(* IEC 61131-3 sources: daoli-st-library/DL_MathData (part 27) *)

(* ---- FC_DL_TrimmedMeanCalc.st ---- *)
(*
  ==================================================================
  组件名 Component  : FC_DL_TrimmedMeanCalc
  分类   Category   : DL_MathData
  前缀   Naming     : FC_DL_ ｜ b/n/u/f/t/e/st 类型前缀制（R265）
  码位   Code ID    : 16#0001_0659 / 065A（故障级）
  版本   Version    : 1.0.0
  复杂度 Complexity  : 中
  功能   Purpose    : 双端截尾均值（稳健统计，抗野点污染的位置估计）：剔除非有限
                      样本后按升序索引对中段区间求均值。
  开源溯源 Origin    : 公开公式 clean-room，参考公开稳健统计教材的双端截尾均值
                      定义（分类与公式借鉴，零代码复制），本件实现、闸门与码位
                      100% 自有。
  许可证 License    : MIT
  参考   Reference  : IEC 61131-3:2013 §6.6 算术运算符；trimmed mean 公开统计定义
  平台   Platform   : 纯 IEC 61131-3（FOR / 四则 / 委托），三平台通用
  依赖   Depends    : FC_DL_SortIndexLReal（索引排序属主，本件委托排序，R140）
  分工声明 Split     : FC_DL_MeanAbsDevCalc（离散度）/ FC_DL_MedianAbsDev（稳健
                      离散度）/ FB_DL_MovingAverage（滑窗均值）互引；本件为双端
                      截尾均值（稳健位置估计），填位置量缺口（R216）。
  归属 Ownership     : 本件无 TYPE 声明；全部引脚为 IEC 标准原生类型。
                      委托件码位随其属主回传（R66）。
  ------------------------------------------------------------------
  边界 Boundary     :
                      一 非有限样本逐条剔除并计入局部 nNonFinite；nNonFinite 口径
                         **不外显**（R62-D7 定稿口径固化），剔除诊断请用
                         FC_DL_SignalStatistics；除子一律用剔除后的 nEff；
                      二 nCount 越域（< 1 或 > 256）或剔净后 nEff = 0 → 故障码
                         0659 早退（除子已证 ≥ 1 才进入均值段）；
                      三 uTrimLo + uTrimHi >= nEff → 组态码 065A 早退（禁把截尾
                         做成空集）；trim 以剔除后有效样本为基准（非入参计数）；
                      四 委托排序返回值与 bValid 由两个独立变量承接后合取
                         （R295 双承接）；委托码随属主回传（R66）；
                      五 均值区间 [uTrimLo, nEff−1−uTrimHi]，除子
                         (nEff − uTrimLo − uTrimHi) ≥ 1 由段 3 闸证明（禁除零）；
                      六 结果复检非有限 → 三件套兜底（R258）；
                      七 纯函数：无记忆量、无定时器、无边沿实例，每调用重算；
                      八 无全局、无外部变量、无物理地址、无指针。
  错误码 Codes      :
    16#0001_0659【故障级】有效样本数越域（nCount < 1 / > 256，或剔净后 nEff = 0）
    16#0001_065A【故障级】截尾组态非法（uTrimLo + uTrimHi >= nEff，截尾成空集）
  码位反证 Note     :
    0659 与 065A 不可合并：前者出口 nEff = 0（无任何有效样本），后者出口 nEff ≥ 1
    （有效样本存在但被截空），nEff 可由输出唯一还原场景（R90）；0659 合并
    「入参越域」与「剔净为空」的理由：两者出口组合完全同形（fMean = 0、nEff = 0、
    bValid = FALSE），按 R90 不另立。
  验收 Acceptance   :
    算法已证（脚本）：未跑 ｜ 编译器已证（三平台）：未跑
    V1 全同样本 + 任意 trim → 均值 = 该值
    V2 trim = 0/0 → 等价普通均值；V3 uTrimLo+uTrimHi = nEff → 码 065A 早退
    V4 nEff − trim = 1（只余 1 个）→ 均值 = 该样本
    V5 nCount = 0 → 码 0659；V6 nCount = 257 → 码 0659 早退
    V7 含 2 个 NaN → nEff 正确缩减（量化断言）
    V8 trim 单端不对称（lo = 2, hi = 0）→ 区间正确
  修订记录 Revision  :
    2026-11-21  v1.0.0  R63 首版（批 2 · 序号 4）
  ==================================================================
*)
FUNCTION FC_DL_TrimmedMeanCalc : BOOL
VAR_IN_OUT
    afSamples : ARRAY[0..255] OF LREAL; // 样本序列 [工程单位]，只读 / the sample series, read only
END_VAR
VAR_INPUT
    nCount  : DINT := 0;    // 有效样本数入参 [个]，合法域 1..256 / the sample count, legal from one to two hundred fifty six
    uTrimLo : USINT := 0;   // 低端截去个数 [个] / the count trimmed from the low end
    uTrimHi : USINT := 0;   // 高端截去个数 [个] / the count trimmed from the high end
END_VAR
VAR_OUTPUT
    fMean   : LREAL := 0.0; // 截尾均值 [工程单位] / the trimmed mean
    nEff    : DINT := 0;    // 参与均值样本数 [个]（剔除非有限后）/ the effective sample count after dropping non finite samples
    bValid  : BOOL := FALSE; // 结果可用 [-] / the result usable flag
    eErr    : UDINT := 16#0000_0000; // 错误码，0 = 正常 / the error code, zero is ok
    bError  : BOOL := FALSE; // 故障标志（故障级码同拍置位，R45 配对）/ the fault flag raised with a fault level code
END_VAR
VAR
    aVal      : ARRAY[0..255] OF LREAL; // 剔除非有限后的有效样本副本 [工程单位] / the finite sample copy
    aIdx      : ARRAY[0..255] OF DINT;  // 委托输出的排序索引排列 [下标] / the sorted permutation from the delegate
    k         : DINT := 0;    // 遍历索引 [下标] / the traversal index
    nNonFinite: DINT := 0;    // 剔除的非有限样本数 [个]（仅局部留档，不外显，R62-D7 口径；诊断请用 FC_DL_SignalStatistics）/ the dropped non finite count, local only and never exposed
    nCountUse : DINT := 0;    // 入参样本数接管量 [个] / the raw input count holder
    nTrim     : DINT := 0;    // 双端截去总数 [个]（升位防 USINT 和溢出）/ the total trimmed count widened before the sum
    nTrimLo   : DINT := 0;    // 低端截去数升位副本 [个] / the low trim count widened
    nTrimHi   : DINT := 0;    // 高端截去数升位副本 [个] / the high trim count widened
    nKeep     : DINT := 0;    // 参与均值样本数（除子）[个] / the kept sample count used as the divisor
    fSum      : LREAL := 0.0; // 区间样本和 [工程单位] / the interval sample sum
    fMeanUse  : LREAL := 0.0; // 均值工作副本 [工程单位] / the working mean copy
    bSortRet  : BOOL := FALSE; // 委托返回值承接量（独立承接，R295）/ the delegate return holder
    bSortValid: BOOL := FALSE; // 委托 bValid 承接量（独立承接，R295）/ the delegate valid holder
    uSortErr  : UDINT := 16#0000_0000; // 委托错误码承接量 [码] / the delegate error code holder
    bSortErr  : BOOL := FALSE; // 委托故障位承接量 / the delegate fault bit holder
    bSortOk   : BOOL := FALSE; // 返回值与可用位合取后的排序可用位 / the conjunction of the return value and the valid flag
END_VAR  // R64 结构补齐：VAR 段缺失的 END_VAR（门禁机械修复）
VAR CONSTANT
    DL_TMC_NMAX  : DINT := 256;      // 样本容量上界 [个]，与数组容量一致 / the capacity aligned with the array
    DL_TMC_ONE   : DINT := 1;        // 整型一常量 [个] / the integer one constant
    DL_TMC_ZERO  : DINT := 0;        // 整型零常量 [个] / the integer zero constant
END_VAR

// 段 1｜返回值与全部出口预置安全值（R45 四段式第一段）/ segment 1, the preset of the return and every outlet
FC_DL_TrimmedMeanCalc := FALSE; // 返回值预置假 / preset the return false
fMean := 0.0; // 均值预置零 [工程单位] / preset the mean zero
nEff := DL_TMC_ZERO; // 有效样本数预置零 [个] / preset the effective count zero
bValid := FALSE; // 可用标志预置假 / preset the validity false
eErr := 16#0000_0000; // 错误码预置正常 / preset the code to ok
bError := FALSE; // 故障标志预置假 / preset the error flag false
nNonFinite := DL_TMC_ZERO; // 剔除计数预置零 [个] / preset the dropped count zero
nCountUse := DL_TMC_ZERO; // 入参计数接管量预置零 [个] / preset the raw count holder zero
nTrim := DL_TMC_ZERO; // 截去总数预置零 [个] / preset the trimmed total zero
nTrimLo := DL_TMC_ZERO; // 低端截去数预置零 [个] / preset the low trim zero
nTrimHi := DL_TMC_ZERO; // 高端截去数预置零 [个] / preset the high trim zero
nKeep := DL_TMC_ZERO; // 除子预置零 [个] / preset the divisor zero
fSum := 0.0; // 区间和预置零 [工程单位] / preset the interval sum zero
fMeanUse := 0.0; // 均值工作副本预置零 [工程单位] / preset the working mean zero
bSortRet := FALSE; // 委托返回值承接量预置假 / preset the delegate return holder false
bSortValid := FALSE; // 委托可用位承接量预置假 / preset the delegate valid holder false
uSortErr := 16#0000_0000; // 委托码承接量预置零 [码] / preset the delegate code zero
bSortErr := FALSE; // 委托故障位承接量预置假 / preset the delegate fault holder false
bSortOk := FALSE; // 排序可用位预置假 / preset the sort usable bit false

// 段 2｜样本数域闸（边界二，早退禁除零）/ segment 2, the sample count domain gate
nCountUse := nCount; // 入参计数接管 [个] / take the raw count
IF (nCountUse < DL_TMC_ONE) OR (nCountUse > DL_TMC_NMAX) THEN // 计数越域 / the count is out of the domain
    eErr := 16#0001_0659; // 故障级：有效样本数越域 / fault grade, the effective sample count is out of the domain
    bError := TRUE; // 同拍置故障标志（R45 配对）/ raise the fault flag on the same scan
    bValid := FALSE; // 结果不可用 / the result is not usable
    RETURN; // 早退 / early return
END_IF

// 段 3｜非有限样本剔除（边界一：除子口径 = 剔除后有效样本数）/ segment 3, drop the non finite samples
FOR k := DL_TMC_ZERO TO nCountUse - DL_TMC_ONE DO // 有界遍历（上界已证 ≤ 256）/ the bounded traversal with a proven ceiling
    IF (afSamples[k] = afSamples[k]) AND ((afSamples[k] - afSamples[k]) = (afSamples[k] - afSamples[k])) THEN // 有限样本 / a finite sample
        aVal[nEff] := afSamples[k]; // 有限样本写入副本 [工程单位] / copy the finite sample
        nEff := nEff + DL_TMC_ONE; // 有效计数推进 [个] / advance the effective count
    ELSE // 非有限样本 / a non finite sample
        nNonFinite := nNonFinite + DL_TMC_ONE; // 剔除计数推进（仅局部留档，不外显）/ advance the dropped count, local only
    END_IF
END_FOR
IF nEff < DL_TMC_ONE THEN // 剔净后无有效样本（与段 2 同码，出口组合不可区分，R90）/ no sample remains after the drop
    eErr := 16#0001_0659; // 故障级：有效样本数越域（此处为剔净后为空）/ fault grade, the effective count is empty after the drop
    bError := TRUE; // 同拍置故障标志（R45 配对）/ raise the fault flag on the same scan
    bValid := FALSE; // 结果不可用 / the result is not usable
    RETURN; // 早退 / early return
END_IF

// 段 4｜截尾组态闸（边界三，trim 以 nEff 为基准；升位防 USINT 和回绕）/ segment 4, the trim configuration gate
nTrimLo := USINT_TO_DINT(uTrimLo); // 低端截去数升位 [个] / widen the low trim count
nTrimHi := USINT_TO_DINT(uTrimHi); // 高端截去数升位 [个] / widen the high trim count
nTrim := nTrimLo + nTrimHi; // 双端总数（DINT 域无回绕）[个] / the trimmed total in the widened domain
IF nTrim >= nEff THEN // 截尾成空集 / the trim leaves an empty set
    eErr := 16#0001_065A; // 故障级：截尾组态非法 / fault grade, the trim configuration is illegal
    bError := TRUE; // 同拍置故障标志（R45 配对）/ raise the fault flag on the same scan
    bValid := FALSE; // 结果不可用 / the result is not usable
    RETURN; // 早退，除子 nKeep 不可为零 / early return, the divisor can never reach zero
END_IF
nKeep := nEff - nTrim; // 参与均值样本数（除子）[个]，已证 ≥ 1 / the kept count, proven at least one

// 段 5｜委托索引排序（R140；返回值与可用位分承后合取，R295）/ segment 5, the delegated index sort
bSortRet := FC_DL_SortIndexLReal(afValues := aVal, nCount := nEff, aIdx => aIdx, bValid => bSortValid, eErr => uSortErr, bError => bSortErr); // 委托排序：两路各自承接 / delegate the sort into two distinct holders
bSortOk := bSortRet AND bSortValid; // 返回值与可用位合取（IEC 未规定两者的求值次序）/ conjoin the two signals since their evaluation order is unspecified
IF (NOT bSortOk) OR bSortErr THEN // 委托失败 / the delegate failed
    eErr := uSortErr; // 委托码回传（码随属主，R66）/ replay the delegate code
    bError := bSortErr; // 委托故障位回传 / replay the delegate fault bit
    bValid := FALSE; // 结果不可用 / the result is not usable
    RETURN; // 早退 / early return
END_IF

// 段 6｜区间求和（索引区间 [uTrimLo, nEff−1−uTrimHi]；除子 nKeep 已证 ≥ 1，边界五）/ segment 6, the interval sum over the trimmed range
FOR k := nTrimLo TO (nEff - DL_TMC_ONE) - nTrimHi DO // 有界遍历中段区间（区间端点已证合法）/ the bounded traversal over the kept range with proven endpoints
    fSum := fSum + aVal[aIdx[k]]; // 区间样本累加 [工程单位] / accumulate the kept samples
END_FOR
fMeanUse := fSum / DINT_TO_LREAL(nKeep); // 截尾均值 = 和 ÷ 参与数 [工程单位]，除子已证 ≥ 1 / the trimmed mean with the proven divisor

// 段 7｜结果复检兜底（三件套，R258）/ segment 7, the result recheck with the three part fallback
IF (fMeanUse <> fMeanUse) OR ((fMeanUse - fMeanUse) <> (fMeanUse - fMeanUse)) THEN // 结果非有限（理论上不可达，防御保留）/ a non finite result, unreachable by theory, kept as a defence
    fMean := 0.0; // 兜底安全值 [工程单位] / the bottom line safe value
    nEff := DL_TMC_ZERO; // 有效数清零（出口与故障场景同形）/ clear the effective count
    eErr := 16#0001_0659; // 故障级：结果非有限（与样本数越域同族一码，出口组合不可区分，R90）/ fault grade under the same family code
    bError := TRUE; // 置故障标志（R45 配对）/ raise the fault flag
    bValid := FALSE; // 结果不可用 / the result is not usable
    RETURN; // 早退 / early return
END_IF

// 段 8｜统一出口 / segment 8, the unified outlet
fMean := fMeanUse; // 均值出口 [工程单位] / the mean outlet
bValid := TRUE; // 结果可用 / the result is usable
FC_DL_TrimmedMeanCalc := TRUE; // 返回成功 / return success
END_FUNCTION

(* ---- FC_DL_TruncEx.st ---- *)
(*
    FC_DL_TruncEx —— 向零取整防御包装（DINT 范围钳位 + NaN 拦截）
    ------------------------------------------------------------------
    分类      : DL_MathData / Math-Round
    前缀      : FC_DL_
    版本      : 1.0.0
    溯源      : IEC 61131-3 标准语义的道莅防御性实现
                （内部委托平台内建函数，外围统一错误码/钳位/双语文档；
                  未复制任何闭源厂商源码，参考实现仅限 MIT/Apache 许可）
    平台      : 纯 IEC 61131-3，CODESYS / TwinCAT / InoProShop 通用
    作者      : 道莅代码库 · PLC编程专家（R15）
    ------------------------------------------------------------------
    功能说明  : 向零取整（委托内建 TRUNC），如 1.9 得 1、-1.9 得 -1。
                NaN 输入拦截返回 0 并置 16#0001_018B；结果超 DINT 范围
                [-2147483648, 2147483647] 时钳位到对应边界并置 16#0001_0259
                （钳位值非真实取整，bValid=FALSE；无穷输入被范围闸自然
                拦截）。先做范围闸再调 TRUNC，保证内建转换永不溢出。
    错误码    : 0000 正常 / 16#0001_018B 入参越界（NaN 已归零） / 16#0001_0259 上溢下溢（已钳位到 DINT 边界）
    修订记录  : 2026-11-16 v1.0.0 首次入库（R15）
*)
FUNCTION FC_DL_TruncEx : DINT
VAR_INPUT
    lrIn : LREAL; // 输入实数 [无量纲]，任意有限值或 NaN/无穷 / input real value [dimensionless], any finite value or NaN/inf
END_VAR
VAR_OUTPUT
    eErr : UDINT; // 错误码，0=正常，1=入参越界，2=上溢下溢 / error id, 0=ok, 1=input out of domain, 2=overflow or underflow
    bError   : BOOL; // 是否出错，eErr 非 0 时为 TRUE / error flag, TRUE when eErr is nonzero
    bValid   : BOOL; // 输出是否有效可用，钳位降级时为 FALSE / output valid, FALSE for clamped degraded results
END_VAR
VAR CONSTANT
    DL_TR_HI : LREAL := 2147483648.0; // DINT 上溢闸 [无量纲]，入参达到即超界 / DINT upper overflow gate [dimensionless]
    DL_TR_LO : LREAL := -2147483649.0; // DINT 下溢闸 [无量纲]，入参达到即超界 / DINT lower overflow gate [dimensionless]
END_VAR

// 段 1｜返回值与错误状态预置，任何早退路径不留脏码 / segment 1, preset return value and error states
FC_DL_TruncEx := 0; // 返回值预置安全值 0 / preset return to safe value 0
eErr      := 16#0000_0000; // 错误码预置正常 / preset error id to ok
bError        := FALSE; // 错误标志预置无错 / preset error flag to FALSE
bValid        := TRUE; // 有效标志预置可用 / preset valid flag to TRUE

// 段 2｜NaN 拦截：自不等判据，归零早退，不进内核 / segment 2, NaN interception by self-inequality, zeroed early exit
IF lrIn <> lrIn THEN
    eErr := 16#0001_018B; // 信息级：输入 NaN，已归零 / informational, NaN input, zeroed
    bError   := TRUE; // 置错误标志 / raise error flag
    bValid   := FALSE; // 输出不可用 / output invalid
    RETURN; // 返回预置安全值 0 / return preset safe value 0
END_IF

// 段 3｜DINT 范围闸：先判后转换，保证内建 TRUNC 永不溢出（无穷输入同样命中闸） / segment 3, DINT range gate, decide before conversion so built-in TRUNC never overflows, infinity hits the gate too
IF lrIn >= DL_TR_HI THEN
    FC_DL_TruncEx := 2147483647; // 上溢钳位到 DINT 上界 / overflow clamped to the DINT upper bound
    eErr      := 16#0001_0259; // 上溢码 / overflow code
    bError        := TRUE; // 置错误标志 / raise error flag
    bValid        := FALSE; // 钳位值非真实取整 / clamped value is not the true truncation
    RETURN;
ELSIF lrIn <= DL_TR_LO THEN
    FC_DL_TruncEx := -2147483648; // 下溢钳位到 DINT 下界 / underflow clamped to the DINT lower bound
    eErr      := 16#0001_0259; // 下溢码 / underflow code
    bError        := TRUE; // 置错误标志 / raise error flag
    bValid        := FALSE; // 钳位值非真实取整 / clamped value is not the true truncation
    RETURN;
END_IF

// 段 4｜域内委托内建 TRUNC（向零取整） / segment 4, in-domain delegation to built-in TRUNC, rounding toward zero
FC_DL_TruncEx := TRUNC(lrIn); // 委托内建 TRUNC 内核，不自实现取整内核 / delegate to built-in TRUNC kernel

// 段 5｜结果复检兜底（防御纵深，正常路径不可达） / segment 5, result recheck as defense in depth
IF (FC_DL_TruncEx <> FC_DL_TruncEx) OR (FC_DL_TruncEx > 2147483647) OR (FC_DL_TruncEx < -2147483648) THEN
    FC_DL_TruncEx := 0; // 兜底安全值 / bottom-line safe value
    IF eErr = 16#0000_0000 THEN
        eErr := 16#0001_018B; // 首事件优先置码 / first-event priority code
        bError   := TRUE; // 置错误标志 / raise error flag
        bValid   := FALSE; // 输出不可用 / output invalid
    END_IF
END_IF
END_FUNCTION

(* ---- FC_DL_TruncToMultipleInt.st ---- *)
(*==============================================================================
 * 组件名称 : FC_DL_TruncToMultipleInt ｜ 子库 : DL_MathData ｜ v1.0.0 ｜ 2026-11-23
 * 平台     : CODESYS 3.5 / TwinCAT 3 / InoProShop / Machine Expert（纯 IEC，无厂商库）
 * 功能简介 : 整数向零截断到 nMultiple 的倍数（丢弃不足一个倍数的余量，
 *            符号随被除数）。纯整数算术实现：整除（ST 中 DIV 对整数
 *            向零截断）后回乘，即得截断对齐结果。
 * 契约     : 返回向零截断结果；nMultiple <= 0 恒返回 0；
 *            纯函数无状态、同输入同输出。
 * 依赖     : 无 DL_ 内部依赖（本批自足实现）
 * 红线自检 : R1 零全局 R2 零%I/%Q R3 纯IEC R4 非法倍数返 0（防除零）
 *            R5 双语注释 R6 N/A（无状态机） R7 N/A（无定时器实例）
 * 修订历史 : 2026-11-23 R78-B1 对齐取整族模板派生首版
 *============================================================================*)
FUNCTION FC_DL_TruncToMultipleInt : DINT
VAR_INPUT
    nValue : DINT;          // 输入整数 / Input integer value
    nMultiple : DINT;       // 对齐倍数，须 > 0 / Alignment multiple, must be > 0
END_VAR
IF nMultiple <= 0 THEN
    FC_DL_TruncToMultipleInt := 0;      // 非法倍数返 0 / Invalid multiple returns 0
    RETURN;
END_IF
FC_DL_TruncToMultipleInt := (nValue / nMultiple) * nMultiple;   // 整除截断回乘 / Truncate by integer division and remultiply
END_FUNCTION

(* ---- FC_DL_UdintToBcd.st ---- *)
(*
    FC_DL_UdintToBcd —— UDINT 到 8 位十进制 BCD 码饱和防御转换
    ------------------------------------------------------------------
    分类      : DL_MathData / Convert
    前缀      : FC_DL_
    版本      : 1.0.0
    溯源      : IEC 61131-3 标准语义的道莅防御性实现
                （内部委托平台内建函数，外围统一错误码/钳位/双语文档；
                  未复制任何闭源厂商源码，参考实现仅限 MIT/Apache 许可）
    平台      : 纯 IEC 61131-3，CODESYS / TwinCAT / InoProShop 通用
    作者      : 道莅代码库 · PLC编程专家（R16）
    ------------------------------------------------------------------
    功能说明  : 将十进制值 nIn（0..99999999）防御性转换为 8 位十进制 BCD 码并返回；
                nIn 超出 99999999 时饱和输出 BCD 码 16#99999999，置信息级 16#0001_01D2
                （与 R9 FC_DL_WordToBcd 的 9999 饱和口径一致，域扩大 4 位）；
                钳位方向：仅上界单侧饱和至 16#99999999；
                域内按除 10 取余逐位拼装半字节：除子为常量 10，编译期恒非零，
                满足除法前判除子非零红线；8 次整除后余数归零，无溢出路径；
                纯整数域输入不存在 NaN/±INF 非有限态，故本组件无故障级路径；
                信息级码属正常防御：bError=FALSE、bValid=TRUE，输出饱和后防御值。
    错误码    : 16#0001_01D2 输入超 99999999，已饱和至 BCD 16#99999999——信息级，正常防御
                16#0001_01D3 预留禁用（信息级，不得挪用）
                16#0001_02A9 预留禁用（故障级，不得挪用）
                16#0001_02AA 预留禁用（故障级，不得挪用）
                16#0001_02AB 预留禁用（故障级，不得挪用）
    状态机    : R6 标注 N/A —— 本组件为纯函数无顺序状态机，无 CASE 可写，非法状态不可能出现，故以本节说明替代 ELSE 兜底
    修订记录  : 2026-11-16 v1.0.0 首次入库（R16）
*)
FUNCTION FC_DL_UdintToBcd : UDINT
VAR_INPUT
    nIn : UDINT; // 十进制值 [0..99999999] / decimal value, 0..99999999
END_VAR
VAR_OUTPUT
    eErr   : UDINT; // 错误码，0=正常 / error id, 0=ok
    bError : BOOL;  // 是否出错，eErr 非 0 时为 TRUE / error flag, TRUE when eErr is nonzero
    bValid : BOOL;  // 输出是否有效可用 / output valid flag
END_VAR
VAR CONSTANT
    DL_BCD8_MAX    : UDINT := 99999999;    // 8 位 BCD 十进制域上界 [无量纲] / 8-digit BCD decimal domain upper bound
    DL_BCD8_SAT    : UDINT := 16#99999999; // 8 位 BCD 饱和输出码（每位半字节 9） [BCD 位] / 8-digit BCD saturating output code (nibble 9 each)
    DL_BCD_NIB_CNT : INT   := 8;           // UDINT 32 位容器 BCD 半字节总数 [个] / total BCD nibble count of 32-bit UDINT container
    DL_DEC_BASE    : UDINT := 10;          // 十进制除法基（编译期常量，恒非零） [基数] / decimal division base (compile-time constant, never zero)
END_VAR
VAR
    i      : INT;   // 半字节循环索引 [个] / nibble loop index
    uDigit : UDINT; // 当前十进制位值（0~9） [位] / current decimal digit value (0~9)
    uTmp   : UDINT; // 剩余待转换商 [无量纲] / remaining quotient to convert
END_VAR

// 段 1｜返回值与错误状态预置 / segment 1, preset return value and error status
FC_DL_UdintToBcd := 0; // 故障缺省返回 0 [BCD 位] / fault default returns 0
eErr   := 0;     // 预置无错误 / preset no error
bError := FALSE; // 预置无故障（整数域无故障态） / preset no fault (no fault states in integer domain)
bValid := FALSE; // 预置无效，通过饱和判定后置位 / preset invalid, set TRUE after saturation check

// 段 2｜上界单侧饱和钳位 / segment 2, upper-bound saturating clamp
IF nIn > DL_BCD8_MAX THEN
    FC_DL_UdintToBcd := DL_BCD8_SAT; // 饱和输出 BCD 16#99999999（与 R9 WordToBcd 口径一致，域扩大 4 位） / saturate to BCD 16#99999999 (aligned with R9 WordToBcd policy, domain widened by 4 digits)
    eErr := 16#0001_01D2;            // 信息级：超上界已饱和 / info level: above upper bound, saturated
    bError := FALSE;                 // 信息级饱和不置故障 / info-level saturation never raises fault
    bValid := TRUE;                  // 饱和输出有效可用 / saturated output is valid
    RETURN;                          // 立即返回 / immediate return
END_IF

// 段 3｜除 10 取余逐位拼装主体计算（末段） / segment 3, divide-by-10 remainder digit assembly main conversion (final)
uTmp := nIn; // 商初始化为输入值 / initialize quotient with input
FOR i := 0 TO DL_BCD_NIB_CNT - 1 DO
    uDigit := uTmp MOD DL_DEC_BASE;       // 除 10 取余得当前十进制位（除子常量 10 恒非零） / modulo 10 for current digit (constant divisor 10, never zero)
    FC_DL_UdintToBcd := FC_DL_UdintToBcd OR SHL(uDigit, 4 * i); // 拼装第 i 个 BCD 半字节（SHL 移位量 4*i ≤ 28 安全） / assemble i-th BCD nibble (shift 4*i <= 28, safe)
    uTmp := uTmp / DL_DEC_BASE;           // 整除 10 前进到下一位（除子常量 10 恒非零） / integer-divide by 10 to next digit (constant divisor 10, never zero)
END_FOR
bError := FALSE; // 域内转换无故障 / in-domain conversion, no fault
bValid := TRUE;  // 输出有效可用 / output valid
END_FUNCTION

(* ---- FC_DL_UdintToDintChk.st ---- *)
(*
    FC_DL_UdintToDintChk —— UDINT 到 DINT 越界钳位防御转换
    ------------------------------------------------------------------
    分类      : DL_MathData / Convert
    前缀      : FC_DL_
    版本      : 1.0.0
    溯源      : IEC 61131-3 标准语义的道莅防御性实现
                （内部委托平台内建函数，外围统一错误码/钳位/双语文档；
                  未复制任何闭源厂商源码，参考实现仅限 MIT/Apache 许可）
    平台      : 纯 IEC 61131-3，CODESYS / TwinCAT / InoProShop 通用
    作者      : 道莅代码库 · PLC编程专家（R16）
    ------------------------------------------------------------------
    功能说明  : 将 UDINT 输入防御性转换为 DINT 并作为返回值输出；
                uIn 超出 DINT 上界 2147483647 时钳位至上界，置信息级 16#0001_01CC；
                钳位方向：仅上界单侧饱和（UDINT 无负值，下界 0 天然落在 DINT 域内无需钳位）；
                纯整数域输入不存在 NaN/±INF 非有限态，亦无除法运算，故本组件无故障级路径；
                域内转换委托平台内建 UDINT_TO_DINT 语义，不重实现数学内核；
                信息级码属正常防御：bError=FALSE、bValid=TRUE，输出钳位后防御值。
    错误码    : 16#0001_01CC 输入超 DINT 上界，已钳位至 2147483647——信息级，正常防御
                16#0001_01CD 预留禁用（信息级，不得挪用）
                16#0001_02A0 预留禁用（故障级，不得挪用）
                16#0001_02A1 预留禁用（故障级，不得挪用）
                16#0001_02A2 预留禁用（故障级，不得挪用）
    状态机    : R6 标注 N/A —— 本组件为纯函数无顺序状态机，无 CASE 可写，非法状态不可能出现，故以本节说明替代 ELSE 兜底
    修订记录  : 2026-11-16 v1.0.0 首次入库（R16）
*)
FUNCTION FC_DL_UdintToDintChk : DINT
VAR_INPUT
    uIn : UDINT; // 待转换输入 [无量纲] / input value to convert
END_VAR
VAR_OUTPUT
    eErr   : UDINT; // 错误码，0=正常 / error id, 0=ok
    bError : BOOL;  // 是否出错，eErr 非 0 时为 TRUE / error flag, TRUE when eErr is nonzero
    bValid : BOOL;  // 输出是否有效可用 / output valid flag
END_VAR
VAR CONSTANT
    DL_DINT32_MAX : UDINT := 2147483647; // DINT 域上界 2147483647 [无量纲] / DINT upper bound 2147483647
END_VAR

// 段 1｜返回值与错误状态预置 / segment 1, preset return value and error status
FC_DL_UdintToDintChk := 0; // 故障缺省返回 0 [无量纲] / fault default returns 0
eErr   := 0;     // 预置无错误 / preset no error
bError := FALSE; // 预置无故障（整数域无故障态） / preset no fault (no fault states in integer domain)
bValid := FALSE; // 预置无效，通过钳位判定后置位 / preset invalid, set TRUE after clamp check

// 段 2｜上界单侧饱和钳位与主体转换（末段） / segment 2, upper-bound saturating clamp and main conversion (final)
IF uIn > DL_DINT32_MAX THEN
    FC_DL_UdintToDintChk := DL_DINT32_MAX; // 正向钳位至 DINT 上界 2147483647 / clamp to DINT upper bound 2147483647
    eErr := 16#0001_01CC;                  // 信息级：超上界已钳位 / info level: above upper bound, clamped
ELSE
    FC_DL_UdintToDintChk := UDINT_TO_DINT(uIn); // 域内委托平台内建 _TO_ 转换语义 / in-domain delegate to built-in _TO_ conversion
    eErr := 0; // 域内无错误 / in-domain, no error
END_IF
bValid := TRUE; // 域内或钳位输出均有效可用 / in-domain or clamped output is valid
END_FUNCTION

(* ---- FC_DL_UdintToLintChk.st ---- *)
(*
    FC_DL_UdintToLintChk —— UDINT 到 LINT 升位验真
    ------------------------------------------------------------------
    分类      : DL_MathData / Convert
    前缀      : FC_DL_
    版本      : 1.0.0
    溯源      : IEC 61131-3 标准语义的道莅防御性实现（UDINT 32 位无符号 → LINT 64 位有符号）；
                委托平台内建 UDINT_TO_LINT 完成升位，本件不重实现数学内核；
                round-trip 验真判据、复核开关、错误分级与码位 100% 自有；
                clean-room 重写，未复制任何闭源厂商源码，参考实现仅限 MIT/Apache 许可
    平台      : 纯 IEC 61131-3，CODESYS V3.5+ / TwinCAT 3 / InoProShop 通用
    作者      : 道莅代码库 · PLC编程专家（R20）
    ------------------------------------------------------------------
    功能说明  : UDINT 到 LINT 在数学上恒无损（32 位无符号域完全落在 64 位有符号域内），
                但平台实现常见两种路径：直接零扩展（正确），或经 32 位有符号中间量再升位
                （错误：≥ 2^31 的值被符号扩展成负数）。后者在 DINT 中转站写法里反复出现，
                且编译期无告警、运行期只在超过 2147483647 时才显形，属隐蔽缺陷。
                本件的价值就是把这个隐性错误变成可判定的显式故障：
                核心防御：① round-trip 验真——把结果 LINT_TO_UDINT 反算回去，
                   与输入逐位相等才算无损；不等即判平台符号扩展错误（故障级）；
                ② 验真是判定式而非猜测式：只依赖 IEC 标准往返转换，不依赖任何平台内建语义；
                ③ bCheckEveryCall = FALSE 时跳过复核以降开销，但发信息级说明
                   「本拍未验真」，让审计侧知道该批数据没有复核保护；
                ④ 反算本身也在域内（LINT 结果必为 0~4294967295，若平台已错则反算必然不等），
                   不存在二次溢出风险。
                职责边界：有符号域内饱和归 FC_DL_LintToDintSat，双向无符号落地归
                FC_DL_LintToUdintSat；本件只承担「升位是否真正无损」的验真职责。
    编译门槛  : 主路径依赖平台内建 UDINT_TO_LINT 与 LINT_TO_UDINT，均为 IEC 61131-3
                标准转换函数，三平台标准库均提供，无厂商方言。
    错误码    : 16#0001_0414 调用方关闭逐次复核（bCheckEveryCall = FALSE），本拍未验真——信息级，值仍可用
                16#0001_0415 预留禁用（信息级，不得挪用）
                16#0001_033C round-trip 验真失败，平台把中间量经 32 位有符号路径符号扩展——故障级，bValid = FALSE
                16#0001_033D 预留（故障级，不得挪用）
                16#0001_033E 预留禁用（故障级，不得挪用）
    码位总账  : 16#0001_0414 用 / 16#0001_0415 预留 ｜ 16#0001_033C 用 / 16#0001_033D 预留 / 16#0001_033E 预留
    状态机    : R6 标注 N/A —— 本组件为纯函数无顺序状态机，无 CASE 可写，非法状态不可能出现
    采样约定  : 本件无定时器、无沿检测、无状态；单拍纯计算，结论与任务周期无关。
                复核开关是引脚量而非内部锁存，调用方可按数据重要性逐调用切换。
    修订记录  : 2026-11-16 v1.0.0 首次入库（R20）
*)
FUNCTION FC_DL_UdintToLintChk : LINT
VAR_INPUT
    uIn              : UDINT;                // 输入值 [无量纲]，全域 0~4294967295 / input value [dimensionless], full UDINT domain
    bCheckEveryCall  : BOOL := TRUE;          // TRUE = 每次调用都做 round-trip 复核 / TRUE performs the round-trip check on every call
END_VAR
VAR_OUTPUT
    eErr             : UDINT;                 // 错误码，0=正常 / error id, 0=ok
    bError           : BOOL;                  // 故障标志，eErr 为故障级时 TRUE / error flag, TRUE on fault-level eErr
    bValid           : BOOL;                  // 返回值是否可用（验真失败为 FALSE）/ return usable, FALSE when the round trip failed
    bRoundTripFail   : BOOL;                  // round-trip 复核失败标志 / round-trip check failed flag
END_VAR
VAR CONSTANT
    DL_UDINT_MAX     : UDINT := 16#FFFF_FFFF; // UDINT 上限值，域上限登记（类型本身即保证无需显式比较）[无量纲] / the UDINT maximum, registered domain top [dimensionless]
    DL_LINT_ZERO     : LINT := 0;             // 有符号零常量，避免裸字面量 [无量纲] / signed zero constant [dimensionless]
END_VAR
VAR
    liOut            : LINT;                  // 升位结果中间量 [无量纲] / widened result intermediate [dimensionless]
    uBack            : UDINT;                 // 反算回无符号的复核值 [无量纲] / back-converted value used by the check [dimensionless]
END_VAR

// 段 1｜返回值与错误状态预置 / segment 1, preset return value and error status
FC_DL_UdintToLintChk := DL_LINT_ZERO;         // 故障缺省返回 0 [无量纲] / fault default returns zero [dimensionless]
eErr := 0;                                    // 预置无错误 / preset no error
bError := FALSE;                              // 预置无故障 / preset no fault
bValid := FALSE;                              // 预置不可用，通过闸门后置位 / preset invalid, set TRUE after the gates
bRoundTripFail := FALSE;                      // 预置未失败 / preset no failure
liOut := DL_LINT_ZERO;                        // 中间量清零 / clear the intermediate

// 段 2｜主体：域内升位委托平台内建（数学上恒无损）/ segment 2, widen through the built-in, mathematically lossless
liOut := UDINT_TO_LINT(uIn);                  // 32 位无符号升 64 位有符号 [无量纲] / widen 32-bit unsigned into 64-bit signed [dimensionless]

// 段 3｜复核开关闸：关闭复核只发信息级，绝不伪装成已验真 / segment 3, check switch gate
IF NOT bCheckEveryCall THEN
    eErr := 16#0001_0414;                     // 信息级：本拍未验真，值仍可用 / info level, unchecked this cycle, still usable
    FC_DL_UdintToLintChk := liOut;            // 发布未复核的结果 / publish the unchecked result
    bValid := TRUE;                           // 未复核不等于不可用 / unchecked does not mean unusable
    RETURN;                                   // 出口 / exit
END_IF

// 段 4｜round-trip 验真：反算回去必须逐位相等 / segment 4, round-trip verification
uBack := LINT_TO_UDINT(liOut);                // 反算回无符号域 [无量纲] / convert back into the unsigned domain [dimensionless]
IF uBack <> uIn THEN
    bRoundTripFail := TRUE;                   // 标记验真失败 / flag the failed verification
    eErr := 16#0001_033C;                     // 故障级：平台符号扩展错误 / fault level, the platform sign-extended the value
    bError := TRUE;                           // 置故障标志 / raise the error flag
    bValid := FALSE;                          // 返回值不可用于后续运算 / the value must not enter later arithmetic
    FC_DL_UdintToLintChk := liOut;            // 仍发布结果供 HMI 对比观察 / still publish the value so HMI can compare it
    RETURN;                                   // 出口 / exit
END_IF

// 段 5｜发布验真通过的结果 / segment 5, publish the verified result
FC_DL_UdintToLintChk := liOut;                // 输出升位结果 [无量纲] / publish the widened result [dimensionless]
bValid := TRUE;                               // 验真通过即可用 / verified values are usable
END_FUNCTION

(* ---- FC_DL_UdintToRealChk.st ---- *)
(*
    FC_DL_UdintToRealChk —— UDINT 到 REAL 精度告警转换
    ------------------------------------------------------------------
    分类      : DL_MathData / Convert
    前缀      : FC_DL_
    版本      : 1.0.0
    溯源      : IEC 61131-3 标准语义的道莅防御性实现
                （接口语义由 IEC 61131-3 定义，内部委托平台内建 UDINT_TO_REAL，
                  外围统一错误码 / 钳位 / 双语文档；clean-room 重写，
                  未复制任何闭源厂商源码，参考实现仅限 MIT/Apache 许可）
    平台      : 纯 IEC 61131-3，CODESYS / TwinCAT / InoProShop 通用
    作者      : 道莅代码库 · PLC编程专家（R17）
    ------------------------------------------------------------------
    功能说明  : 将 UDINT 防御性转换为 REAL 并作为返回值输出，转换委托平台内建 UDINT_TO_REAL；
                nIn 超过 2^24（16777216，REAL 尾数 24 位可精确表示的整数上界）时，
                值照常转换输出，仅置信息级 16#0001_01FE 提示低位精度损失（bError=FALSE、bValid=TRUE）；
                负值分支结构性不存在（UDINT 为无符号类型，由类型系统保证），故无下界比较；
                本件只对 REAL 目标域立项：UDINT 全域 ≤ 2^32 远小于 2^53，转 LREAL 恒无损，
                故不设 UDINT 到 LREAL 的告警件（该结论在此声明，后续轮次不得重复立项）；
                钳位方向：无钳位（信息级仅记录，转换结果为最接近的可表值）。
    错误码    : 16#0001_01FE nIn 超 2^24 精度极限，转换值低位可能失真——信息级，正常防御
                16#0001_01FF 预留禁用（信息级，不得挪用）
                16#0001_02EB 预留禁用（故障级，不得挪用）
                16#0001_02EC 预留禁用（故障级，不得挪用）
                16#0001_02ED 预留禁用（故障级，不得挪用）
    状态机    : R6 标注 N/A —— 本组件为纯函数无顺序状态机，无 CASE 可写，非法状态不可能出现，故以本节说明替代 ELSE 兜底
    修订记录  : 2026-11-16 v1.0.0 首次入库（R17）
*)
FUNCTION FC_DL_UdintToRealChk : REAL
VAR_INPUT
    nIn : UDINT; // 待转换无符号整数值，建议域 0 ~ 4294967295 [无量纲] / unsigned integer to convert, suggested domain 0 .. 4294967295 [dimensionless]
END_VAR
VAR_OUTPUT
    eErr   : UDINT; // 错误码，0=正常 / error id, 0=ok
    bError : BOOL;  // 是否出错，eErr 非 0 时为 TRUE / error flag, TRUE when eErr is nonzero
    bValid : BOOL;  // 输出是否有效可用 / output valid flag
END_VAR
VAR CONSTANT
    DL_F24_MAX_U : UDINT := 16777216; // REAL 尾数 24 位可精确表示的无符号整数上界 2^24 [无量纲] / 2^24 exact-integer bound of REAL's 24-bit significand [dimensionless]
    DL_REAL_ZERO : REAL  := 0.0;      // 返回值预置零（本件无故障路径，仅作预置约定） [无量纲] / preset zero, no fault path in this component [dimensionless]
END_VAR

// 段 1｜返回值与错误状态预置 / segment 1, preset return value and error status
FC_DL_UdintToRealChk := DL_REAL_ZERO; // 预置 0.0（本件无故障级路径，仅作预置约定） [无量纲] / preset 0.0, no fault-level path in this component [dimensionless]
eErr   := 0;     // 预置无错误 / preset no error
bError := FALSE; // 预置无故障（本件无故障级路径） / preset no fault, no fault-level path here
bValid := FALSE; // 预置输出无效，通过精度判定后置位 / preset invalid, set TRUE after the precision check

// 段 2｜24 位尾数精度极限判定与主体转换（末段） / segment 2, 24-bit significand precision check and main conversion (final)
FC_DL_UdintToRealChk := UDINT_TO_REAL(nIn); // 值照常转换（委托平台内建转换语义），本件只告警不钳位 [无量纲] / convert as-is via the built-in conversion, this component warns but never clamps [dimensionless]
IF nIn > DL_F24_MAX_U THEN // 无符号类型仅需上界单侧比较，负值分支由类型系统结构性排除 [无量纲] / unsigned type only needs the upper-bound test, negative branch excluded by the type system [dimensionless]
    eErr := 16#0001_01FE; // 信息级：超 2^24 精度极限，低位可能失真，仅记录不钳位 / info level: beyond the 2^24 precision limit, low bits may lose accuracy, recorded only
ELSE
    eErr := 0;            // 精度域内无告警 / within the precision domain, no notice
END_IF
bError := FALSE; // 信息级精度告警不置故障 / info-level precision notice never raises fault
bValid := TRUE;  // 域内或精度告警输出均有效可用 / in-domain or precision-noticed output is valid
END_FUNCTION

(* ---- FC_DL_UdintToStringTrim.st ---- *)
(*
    FC_DL_UdintToStringTrim —— UDINT 到定宽十进制字段（右对齐）的防御字符串化
    ------------------------------------------------------------------
    分类      : DL_MathData / Convert
    前缀      : FC_DL_
    版本      : 1.0.0
    溯源      : IEC 61131-3 标准语义的道莅防御性实现（UDINT → STRING 定宽右对齐补位，
                委托平台内建 UDINT_TO_STRING 与标准串函数 LEN / LEFT / CONCAT；
                补位、四步截断样板、目标宽度闸、错误分级与码位 100% 自有；
                clean-room 编写，未复制任何闭源厂商源码）
    平台      : 纯 IEC 61131-3，CODESYS 3.5 / TwinCAT 3 / InoProShop / Machine Expert 通用
    作者      : 道莅代码库 · PLC编程专家（R69 构建轮 · 批 1 · N3）
    ------------------------------------------------------------------
    功能说明  : R22 定宽字段族的无符号补口。库内已有 FC_DL_DintToStringTrim（有符号，
                去前导空格左对齐）与 FC_DL_LrealToStringTrim（浮点）——本件补 UDINT
                方向，且语义与有符号版**异构**，不可互相替代：
                ① 有符号版做「修剪」（去掉平台补的前导空格后左对齐）；
                   本件做「定宽右对齐」（按目标宽度左补空格，供报表 / 报文定宽字段）。
                ② 上界语义异构：DINT 上界 2147483647 为 10 位数，UDINT 上界
                   4294967295 为 10 位数但**多一个符号位宽**——若把 UDINT 值先转 DINT
                   （现场常见写法），大于 2147483647 的值会翻成负数并输出「-294967296」
                   ！本件全程在 UDINT 域内字符串化，禁止任何有符号中转（R55/R56 口径：
                   浮点 / 有符号 → 无符号必须双分支显式，此处根本不做中转）。
                ③ 目标宽度 uFieldWidth 域 1..32：0 宽度无意义（故障级）；超 32 亦为故障级
                   ——补位源是 32 字符空格常量，宽度超过补位源时 LEFT 会静默返回全长，
                   表现为「字段比要求窄」，故必须在域闸挡住而不得靠钳位；
                   宽度小于实际位数且 bAllowTrunc = FALSE 时返回空串并报故障级，
                   绝不返回半截数值（把 4294967295 写成 429 上位机会当真数据）。
                补位实现：用常量空格串 + LEFT 取 nPad 个 + CONCAT 前缀，禁 WHILE 拼串
                （拼串随长度平方级增长，且串函数异常时会死循环）。
    错误码    : 16#0001_04F8 已按目标宽度左补空格（bPadded 可查）—— 信息级，值可用
                16#0001_04F9 发生截断且 bAllowTrunc = TRUE（bTruncated 可查）—— 信息级，值可用
                16#0001_03FA 目标宽度非法（uFieldWidth = 0）—— 故障级，返回空串
                16#0001_03FB 需要截断但 bAllowTrunc = FALSE —— 故障级，返回空串
    码位总账  : 16#0001_03FA / 03FB 用 ｜ 16#0001_04F8 / 04F9 用
    状态机    : R6 标注 N/A —— 纯函数无顺序状态机，无 CASE 可写，非法状态不可能出现
    采样约定  : 无定时器 / 无沿检测 / 无跨周期状态，结论与任务周期无关
    修订记录  : 2026-11-22 v1.0.0 首次入库（R69 构建轮 · 批 1 · N3）
*)
FUNCTION FC_DL_UdintToStringTrim : STRING(255)
VAR_INPUT
    uIn          : UDINT;                      // 待字符串化的无符号值 [无量纲]，全域 0..4294967295 / unsigned value, full UDINT domain
    uFieldWidth  : USINT := 10;                // 定宽字段宽度 [字符]，域 1..32 / fixed field width [characters], 1 to 32
    bAllowTrunc  : BOOL := FALSE;              // TRUE = 允许截断；FALSE = 需截断即故障 / TRUE allows truncation
END_VAR
VAR_OUTPUT
    eErr         : UDINT;                      // 错误码，0 = 正常 / error id, 0 = ok
    bError       : BOOL;                       // 故障标志，故障级码时为 TRUE / error flag, TRUE on fault level
    bValid       : BOOL;                       // 返回值是否可用（故障级为 FALSE）/ return usable, FALSE on fault level
    bPadded      : BOOL;                       // 本次做了左补空格 / left padding happened
    bTruncated   : BOOL;                       // 本次发生截断 / truncation happened
END_VAR
VAR CONSTANT
    DL_US_CAP    : INT := 255;                 // STRING 型长度上限 [字符]（R49 口径）/ STRING capacity [characters]
    DL_US_W_MIN  : USINT := 1;                 // 目标宽度下限 [字符] / field width floor [characters]
    DL_US_W_MAX  : INT := 32;                  // 目标宽度上限 [字符]，等于补位源空格串长度（超此宽度补位不可信）/ width ceiling [characters]
    DL_US_BLANKS : STRING(32) := '                                ';  // 32 个空格常量，补位源 [字符] / 32 blanks, the padding source
    DL_US_EMPTY  : STRING(1) := '';            // 空串常量，故障缺省返回 / empty string returned on faults
    DL_US_ZERO   : INT := 0;                   // 整型零常量，避免裸字面量 [字符] / integer zero constant
END_VAR
VAR
    sRaw         : STRING(255);                // 内建字符串化原始结果 / raw result of the built-in conversion
    sPad         : STRING(32);                 // 左补空格串 / left padding string
    sOut         : STRING(255);                // 最终输出串 / final output string
    nLen         : INT;                        // 原始串有效长度，一次锁存 [字符] / latched raw length [characters]
    nWidth       : INT;                        // 目标宽度，由引脚转出 [字符] / target width from the pin [characters]
    nPad         : INT;                        // 需要补的空格个数 [字符] / number of blanks to add
END_VAR

// 段 1｜返回值与错误状态预置（实战规则 1①）/ segment 1, preset the return value and the status
FC_DL_UdintToStringTrim := DL_US_EMPTY;   // 故障缺省返回空串 / fault default returns an empty string
eErr       := 0;                          // 预置无错误 / preset no error
bError     := FALSE;                      // 预置无故障 / preset no fault
bValid     := FALSE;                      // 预置不可用 / preset unusable
bPadded    := FALSE;                      // 预置未补位 / preset unpadded
bTruncated := FALSE;                      // 预置未截断 / preset untruncated

// 段 2｜目标宽度闸：0 宽度无意义，先判后算 / segment 2, field width gate
IF uFieldWidth < DL_US_W_MIN THEN
    eErr   := 16#0001_03FA;               // 故障级：目标宽度非法 / fault level: illegal field width
    bError := TRUE;                       // R45 配对 / paired with the code
    bValid := FALSE;                      // 返回值不可用 / return unusable
    RETURN;                               // 出口，不触碰内建 / exit, the built-in is never touched
END_IF
nWidth := USINT_TO_INT(uFieldWidth);      // 宽度转整型 [字符] / width to INT [characters]
IF nWidth > DL_US_W_MAX THEN
    eErr   := 16#0001_03FA;               // 故障级：宽度超补位源上限（32），补位不可信 / fault level: width above the padding source
    bError := TRUE;                       // R45 配对 / paired with the code
    bValid := FALSE;                      // 返回值不可用 / return unusable
    RETURN;                               // 出口 / exit
END_IF

// 段 3｜主体：委托平台内建字符串化（全程无有符号中转）/ segment 3, delegate the built-in in the unsigned domain
sRaw := UDINT_TO_STRING(uIn);             // 无符号值 → 原始串，绝不先转 DINT（反例会输出负数）/ unsigned to string, never via DINT
nLen := LEN(sRaw);                        // 原始串长度，一次锁存 [字符] / latch the size exactly once [characters]
IF nLen > DL_US_CAP THEN
    nLen := DL_US_CAP;                    // 超容量按上限钳位 [字符] / clamp to the capacity [characters]
ELSIF nLen < DL_US_ZERO THEN
    nLen := DL_US_ZERO;                   // 负长度防御，结构性不可达 [字符] / negative length guard, unreachable
END_IF

// 段 4｜四步截断样板（R37）：长度已锁存 → 宽度比较 → 标志先置 → 按允许分路
// segment 4, the four-step truncation pattern: latch, compare, flag first, then branch
IF nLen > nWidth THEN
    bTruncated := TRUE;                   // 标志先于任何写入 / the flag precedes every write
    IF bAllowTrunc THEN
        sOut := LEFT(sRaw, nWidth);       // 允许截断：按宽度截取 / truncation allowed, take the width
        eErr := 16#0001_04F9;             // 信息级：发生截断，值可用 / info level: truncated, still usable
    ELSE
        eErr   := 16#0001_03FB;           // 故障级：需截断但未允许 / fault level: truncation needed but not allowed
        bError := TRUE;                   // R45 配对 / paired with the code
        bValid := FALSE;                  // 返回值不可用 / return unusable
        FC_DL_UdintToStringTrim := DL_US_EMPTY;   // 返回空串，绝不返回半截数值 / never a partial number
        RETURN;                           // 出口 / exit
    END_IF
ELSE
    // 段 5｜右对齐补位：nPad = 宽度 − 位数，LEFT 取空格 + CONCAT 前缀 / segment 5, right-align padding
    nPad := nWidth - nLen;                // 需要补的空格数 [字符] / blanks to add [characters]
    IF nPad > DL_US_ZERO THEN
        sPad := LEFT(DL_US_BLANKS, nPad); // 取 nPad 个空格（禁 WHILE 拼串）/ take the blanks with LEFT
        sOut := CONCAT(sPad, sRaw);       // 空格前缀 + 原始串 = 定宽右对齐 / padding plus the raw string
        bPadded := TRUE;                  // 补位发生 / padding happened
        eErr    := 16#0001_04F8;          // 信息级：已按宽度左补空格 / info level: left padded to the width
    ELSE
        sOut := sRaw;                     // 位数恰等于宽度：直通，无码 / exactly the width, no code
    END_IF
END_IF

// 段 6｜发布结果 / segment 6, publish the result
FC_DL_UdintToStringTrim := sOut;          // 输出最终串 / publish the final string
bValid := TRUE;                           // 补位 / 截断 / 直通三条路径均可用 / usable in every published path
bError := FALSE;                          // 信息级不置故障（双保险）/ info level never raises a fault
END_FUNCTION

(* ---- FC_DL_WeekNumIsoCalc.st ---- *)
(*
  ==================================================================
  组件名 Component  : FC_DL_WeekNumIsoCalc
  分类   Category   : DL_MathData
  版本   Version    : 1.0.0
  功能   Purpose    : ISO 8601 周号计算：输入公历日期，输出 ISO 周号（1~53）
                      与 ISO 周年。全整数实现「儒略日偏移法」：先折儒略日数
                      JDN（整数式，全程正数域整除=向下取整，无符号陷阱），
                      再由「本周四的 JDN」定位所属 ISO 周年，最后以
                      「周年首个周四」为基准做整除求周号。禁 TRUNC 技巧、
                      禁浮点参与，逐整数分支推导。
  来源   Source     : t2-1-lgf-dateandtimer（日期族：JDN 整数式为公开历法
                      口径（Richards 算法公开条款），实现零源码复制）
  互引   Cross-ref  : FC_DL_DayOfWeekCalc（同族星期原子，本件内部 wd 计算
                      与其同口径：JDN mod 7，0=周一）；FC_DL_LeapYearChk
                      （闰年判据同口径，本件以本地常量实现同口径逻辑）
  平台   Platform   : 纯 IEC 61131-3 整数四则 + MOD，三平台通用
  依赖   Depends    : 无 DL_ 内部依赖；无标准库
  归属   Ownership  : 闰年判定以本地常量实现，判据与 FC_DL_LeapYearChk 严格
                      同口径：(y mod 4 = 0 且 y mod 100 <> 0) 或 y mod 400 = 0；
                      本件不声明新枚举。
  红线   Redline    : R1 零全局/VAR_EXTERNAL/R2 零 %I/%Q/R3 纯 IEC 标准
                      R4 月/日域闸 + 年域闸 + 除数全为正常量（结构性无除零）
                      R5 全变量双语同行注释/R6 纯函数无状态机（CASE 不适用）
                      R7 无定时器与沿检测/R8 域界与容差全常量化
  错误码 Codes      : 01【失效级】非法日期（月 1~12 / 日 1~当月天数外）
                      02【失效级】年份域外（有效域 1990~2100）
  码位反证 Note     : 01 与 02 分立依据（R90）：01 在「域内年份 + 日期非法」
                      可观测、02 在「年份域外」可观测，两输入面不同；
                      bValid/nErrId 双通道可区分，无第三码需求。
  验收   Acceptance : V1 2026-11-22（周日）→ 周 47 / 周年 2026 ｜
                      V2 2026-01-01（周四）→ 周 1 / 2026 ｜
                      V3 2026-12-28（周一，周四落 2027）→ 周 53 / 周年 2026
                      ｜ V4 2027-01-01 → 周年 2026 周 53 ｜ V5 2 月 30 → 码 01
                      ｜ V6 1989 或 2101 → 码 02 ｜ V7 2024-02-29（闰）合法
  变更   Revision   : 2026-11-22  v1.0.0  R66 首版（编码阶段批 1 序 4）
  ==================================================================
*)
FUNCTION FC_DL_WeekNumIsoCalc : UINT
VAR_INPUT
    nYear    : UINT;  // 公历年 [年]，有效域 1990~2100 / the calendar year, valid 1990 to 2100
    nMonth   : UINT;  // 公历月 [月]，有效域 1~12 / the calendar month, valid 1 to 12
    nDay     : UINT;  // 公历日 [日]，有效域 1~当月天数 / the calendar day, valid 1 to days in month
END_VAR
VAR_OUTPUT
    nIsoWeek : UINT;  // ISO 周号 1~53 [周] / the ISO week number [week]
    nIsoYear : UINT;  // ISO 周年 [年]（含跨年周归属）/ the ISO week year with cross year attribution
    bValid   : BOOL;  // 结果可用标志 [-] / the result usable flag
    nErrId   : UDINT; // 错误码，0=正常，01=非法日期，02=年域外 [码] / the error code [code]
END_VAR
VAR
    y        : DINT;  // 年工作寄存器 [年] / the year working register
    m        : DINT;  // 月工作寄存器 [月] / the month working register
    d        : DINT;  // 日工作寄存器 [日] / the day working register
    bLeap    : BOOL;  // 闰年判定结果（与 FC_DL_LeapYearChk 同口径）[-] / the leap year verdict, same criteria as the family checker
    uDim     : DINT;  // 当月天数 [日] / the days in the current month
    a        : DINT;  // JDN 折算中间量 (14-m)/12 / the JDN intermediate (14 minus m) over 12
    y2       : DINT;  // JDN 折算年中间量 / the JDN shifted year
    m2       : DINT;  // JDN 折算月中间量 / the JDN shifted month
    jdn      : DINT;  // 输入日期儒略日数 [日] / the Julian day number of the input date
    wd       : DINT;  // 星期序号 0=周一..6=周日 [日] / the weekday index, zero is Monday
    jThu     : DINT;  // 本周周四的 JDN [日] / the JDN of this week's Thursday
    jJanY    : DINT;  // 输入年 1 月 1 日 JDN [日] / the JDN of the input year's Jan 1
    jJanPrev : DINT;  // 前一年 1 月 1 日 JDN [日] / the JDN of the previous year's Jan 1
    jJanNext : DINT;  // 次年 1 月 1 日 JDN [日] / the JDN of the next year's Jan 1
    isoY     : DINT;  // ISO 周年工作寄存器 [年] / the ISO week year working register
    jRef     : DINT;  // ISO 周年 1 月 1 日 JDN [日] / the JDN of the ISO year's Jan 1
    wd0101   : DINT;  // ISO 周年元旦星期序号 [日] / the weekday of the ISO year's Jan 1
    off      : DINT;  // 元素距首个周四的偏移 [日] / the offset from Jan 1 to the first Thursday
    jThu1    : DINT;  // ISO 周年首个周四 JDN [日] / the JDN of the ISO year's first Thursday
    nWeek    : DINT;  // 周号工作寄存器 [周] / the week number working register
END_VAR
VAR CONSTANT
    WIC_Y_MIN    : DINT := 1990;           // 年份有效域下限 [年] / the valid year lower bound
    WIC_Y_MAX    : DINT := 2100;           // 年份有效域上限 [年] / the valid year upper bound
    WIC_JDN_1970 : DINT := 2440588;        // JDN 基准锚点（1970-01-01，星期四）[日] / the JDN anchor of 1970-01-01, a Thursday
    WIC_ERR_NONE  : UDINT := 16#0000_0000; // 无错误 [码] / no error [code]
    WIC_ERR_DATE  : UDINT := 16#0000_0001; // 码 01：非法日期 / code 01, illegal date
    WIC_ERR_YEAR  : UDINT := 16#0000_0002; // 码 02：年域外 / code 02, year out of domain
END_VAR

// 段 1｜输出预置 / segment 1, preset the outputs
FC_DL_WeekNumIsoCalc := UINT#0;  // 失效缺省返回 0 / fault default returns zero
nIsoWeek := UINT#0;              // 周号预置 0 / preset the week to zero
nIsoYear := UINT#0;              // 周年预置 0 / preset the week year to zero
bValid   := FALSE;               // 预置不可用 / preset unusable
nErrId   := WIC_ERR_NONE;        // 预置无错误 / preset no error

// 段 2｜年份域闸（码 02，结构 RETURN 早退）/ segment 2, the year domain gate
IF (nYear < UINT#1990) OR (nYear > UINT#2100) THEN        // 域外年份 / year outside the domain
    nErrId := WIC_ERR_YEAR;
    RETURN;
END_IF

// 段 3｜月/日域闸 + 当月天数（闰年本地常量实现，与 FC_DL_LeapYearChk 同口径）
//      segment 3, month and day gates with the local days in month table
y := UINT_TO_DINT(nYear);       // 年入工作寄存器 / move the year into the register
m := UINT_TO_DINT(nMonth);      // 月入工作寄存器 / move the month into the register
d := UINT_TO_DINT(nDay);        // 日入工作寄存器 / move the day into the register
IF (m < 1) OR (m > 12) THEN     // 月域闸（码 01）/ the month gate, code 01
    nErrId := WIC_ERR_DATE;
    RETURN;
END_IF
bLeap := ((y MOD 4 = 0) AND (y MOD 100 <> 0)) OR (y MOD 400 = 0);  // 闰年判据（同口径）/ the leap criteria, family aligned
CASE m OF        // 当月天数表 / the days in month table
1, 3, 5, 7, 8, 10, 12:  uDim := 31;   // 大月 / the long months
4, 6, 9, 11:            uDim := 30;   // 小月 / the short months
2:                      IF bLeap THEN uDim := 29; ELSE uDim := 28; END_IF  // 二月按闰年 / February by leap
ELSE                    uDim := 0;    // CASE 兜底（结构性不可达，月域已闸）/ unreachable else, the month is gated
END_CASE
IF (d < 1) OR (d > uDim) THEN   // 日域闸（码 01）/ the day gate, code 01
    nErrId := WIC_ERR_DATE;
    RETURN;
END_IF

// 段 4｜JDN 整数折算（Richards 公开式，全程正数域，整除=向下取整）
//      segment 4, the integer JDN conversion, all positive so truncation is floor
a  := (14 - m) DIV 12;                   // m≥1 保证 14-m ≥ 2，商为 0 或 1 / the month shift term
y2 := y + 4800 - a;                      // 折算年，约 6800 量级，DINT 安全 / the shifted year
m2 := m + 12 * a - 3;                    // 折算月 0~11 / the shifted month
jdn := d + (153 * m2 + 2) DIV 5 + 365 * y2 + y2 DIV 4 - y2 DIV 100 + y2 DIV 400 - 32045;  // 儒略日数 [日] / the Julian day number
IF (jdn < WIC_JDN_1970) THEN             // 防御性锚点闸（域内年份结构上不可能触发，留档）/ defensive anchor gate, unreachable in domain
    nErrId := WIC_ERR_YEAR;
    RETURN;
END_IF

// 段 5｜星期与本周四：JDN mod 7 得 0=周一..6=周日（与 FC_DL_DayOfWeekCalc 同口径）
//      segment 5, the weekday and this week's Thursday, family aligned weekday rule
wd   := jdn MOD 7;                       // 星期序号 / the weekday index
jThu := jdn + 3 - wd;                    // 本周周四（wd=3 即周四自身）/ the Thursday of this week

// 段 6｜ISO 周年归属：本周四落在哪个公历年即归属该年
//      segment 6, the ISO year attribution by where this week's Thursday falls
//      三个元旦 JDN 用「本年元旦 ± 365/366」等差推算（闰差由闰年判据决定），
//      不引入辅助 POU，保持单文件自洽：
//      the three Jan 1 JDNs are derived arithmetically, no helper POU, single file self contained
jJanY    := 1 + (153 * 10 + 2) DIV 5 + 365 * (y + 4800 - 1) + (y + 4800 - 1) DIV 4
            - (y + 4800 - 1) DIV 100 + (y + 4800 - 1) DIV 400 - 32045;
            // 本年元旦 JDN（1 月：a=1, m2=10, d=1 代入段 4 同式）/ this year Jan 1 JDN, month terms substituted
bLeap    := ((y MOD 4 = 0) AND (y MOD 100 <> 0)) OR (y MOD 400 = 0);          // 本年闰否 [-] / this year leap flag
IF bLeap THEN
    jJanNext := jJanY + 366;             // 本年为闰 → 次年元旦 = 本年元旦 + 366 / the next Jan 1 is 366 days ahead
ELSE
    jJanNext := jJanY + 365;             // 平年 365 / 365 in a common year
END_IF
IF ((y - 1) MOD 4 = 0) AND NOT (((y - 1) MOD 100 = 0) AND ((y - 1) MOD 400 <> 0)) THEN
    jJanPrev := jJanY - 366;             // 前年为闰 → 本年元旦 = 前年元旦 + 366 / the previous year was leap
ELSE
    jJanPrev := jJanY - 365;             // 前年平年 / the previous year was common
END_IF
IF jThu >= jJanNext THEN                 // 周四落次年 → 归次年 / the Thursday in the next year
    isoY := y + 1;
    jRef := jJanNext;
ELSIF jThu >= jJanY THEN                 // 周四落本年 → 归本年 / the Thursday in this year
    isoY := y;
    jRef := jJanY;
ELSE                                     // 周四落前年 → 归前年 / the Thursday in the previous year
    isoY := y - 1;
    jRef := jJanPrev;
END_IF

// 段 7｜ISO 周年首个周四：从元旦起找第一个 wd=3（周四）
//      segment 7, the ISO year's first Thursday from its Jan 1
wd0101 := jRef MOD 7;                    // 元旦星期序号 / the Jan 1 weekday
IF wd0101 <= 3 THEN
    off := 3 - wd0101;                   // 周四在本周内，向前推 / the Thursday is inside this week
ELSE
    off := 10 - wd0101;                  // 周四在下一周，跨周推 / the Thursday falls into the next week
END_IF
jThu1 := jRef + off;                     // 首个周四 JDN / the first Thursday JDN

// 段 8｜周号整除求解：两周四之差恒为 7 的倍数，DIV 无余数陷阱
//      segment 8, the week number by exact division of two Thursdays
nWeek := (jThu - jThu1) DIV 7 + 1;       // 周号 1~53 [周] / the week number, 1 to 53
IF (nWeek < 1) OR (nWeek > 53) THEN      // 防御性输出域闸（整数法结构上不越域，留档）/ defensive output domain gate
    nErrId := WIC_ERR_DATE;
    RETURN;
END_IF

// 段 9｜出口（ISO 周年归属逻辑上恒在 1989~2101，转 UINT 安全）
//      segment 9, exit, the ISO year stays inside the UINT safe range by construction
nIsoWeek := DINT_TO_UINT(nWeek);         // 发布周号 / publish the week number
nIsoYear := DINT_TO_UINT(isoY);          // 发布周年 / publish the week year
bValid   := TRUE;                        // 结果可用 / the result is usable
FC_DL_WeekNumIsoCalc := nIsoWeek;        // 返回值与输出同源（R191 名实双出口）/ the return mirrors the output
END_FUNCTION

(* ---- FC_DL_WeightedMeanCalc.st ---- *)
(*
  FC_DL_WeightedMeanCalc  —  数组加权平均（权重和防零） / Weighted mean over arrays with zero-sum guard
  分类 Category : DL_MathData
  版本 Version  : 1.0.0
  来源 Source   : t2-1-lgf-math — 统计底座族零检索深化
  溯源 Origin   : clean-room 实现，未复制任何源码行
  功能 Function : 1) 对前 nCnt 个元素计算 SUM(aVals[i] × aWeights[i]) / SUM(aWeights[i])；
                  2) LREAL 域累加；权重和 <= 0 或非有限 → 防除零拒绝，返回 0 + 故障级 03E1；
                  3) 非有限样本/权重元素跳过（不计入累加），剔除后仍有有效元素则正常出值
                  并置信息级 04A4；
                  4) nCnt <= 0 或越界（> 32）先行判界拒绝。
  边界 Boundary : ① 判界先行：nCnt 域检查在累加前完成，越界直接故障出口；
                  ② 除零防御：分母 fWSum 与 DL_WMC_TOL 比较后才做除法；
                  ③ 非有限判定用自反判（x <> x），禁近似阈值；
                  ④ 无 GVL 依赖：纯函数，无外部变量引用，无物理 IO 地址。
  依赖 Depends  : 仅 Standard.library（ABS / LREAL 算术）
  码表 Error codes（段 0001，窗口 03E1 / 04A4）:
    16#0001_03E1 故障级：入参非法（nCnt <= 0 或 > 32，或有效权重和 <= 0 防除零拒绝），
                 返回 0，bValid = FALSE，bError = TRUE
    16#0001_04A4 信息级：非有限元素已剔除（剔除后仍有效，结果照常输出）
  修订历史 Revision :
    2026-11-19  v1.0.0  R41 首版（批次 1 · 序号 4）
*)

FUNCTION FC_DL_WeightedMeanCalc : LREAL
VAR_INPUT
    aVals       : ARRAY[1..32] OF LREAL;   // 样本数组 [EU]，前 nCnt 个参与 / Sample array, first nCnt used
    aWeights    : ARRAY[1..32] OF LREAL;   // 权重数组 [无量纲]，与样本一一对应 / Weight array, one per sample
    nCnt        : INT;               // 参与元素数 [个]，域 1..32 / Element count, 1..32
END_VAR
VAR_OUTPUT
    eErr        : UDINT;             // 事件码，0 = 正常 / Event code
    bError      : BOOL;              // 故障级标志 / Fault-level flag
    bValid      : BOOL;              // 返回值是否可用 / Result usable flag
END_VAR
VAR
    nGuard      : INT;               // 循环守卫计数 [次] / Loop guard counter
    i           : INT;               // 循环游标 [索引] / Loop cursor
    fNum        : LREAL;             // 分子累加器 [EU·权] / Numerator accumulator
    fWSum       : LREAL;             // 分母权重和累加器 [无量纲] / Denominator weight accumulator
    bSkipped    : BOOL;              // 非有限元素剔除标志 / Non-finite element skipped flag
END_VAR
VAR CONSTANT
    DL_WMC_N_MAX     : INT := 32;               // 数组容量上限 [个] / Array capacity bound
    DL_WMC_GUARD_MAX : INT := 32;               // 守卫上限（须 >= N_MAX）/ Loop guard bound
    DL_WMC_TOL       : LREAL := 1.0E-12;        // 权重和有效阈 [无量纲] / Weight-sum validity threshold
    DL_WMC_ERR_IN    : UDINT := 16#0001_03E1;   // 故障级：入参非法 / Fault: invalid input
    DL_WMC_INFO_SKIP : UDINT := 16#0001_04A4;   // 信息级：非有限剔除 / Info: non-finite skipped
END_VAR

(* —— 段 1｜返回值与错误状态预置 —— *)
FC_DL_WeightedMeanCalc := 0.0;      // 缺省返回 0 / default return zero
eErr := 16#0000_0000;               // 预置无事件 / preset no event
bError := FALSE;                    // 预置无故障 / preset no fault
bValid := FALSE;                    // 预置不可用 / preset unusable
fNum := 0.0;                        // 分子清零 / clear numerator
fWSum := 0.0;                       // 分母清零 / clear denominator
bSkipped := FALSE;                  // 剔除标志清零 / clear skip flag
nGuard := 0;                        // 守卫清零（FC 局部量每次调用须显式初始化）/ clear guard
i := 0;                             // 游标清零 / clear cursor

(* —— 段 2｜判界先行：nCnt 域闸（越界直接故障出口） —— *)
IF (nCnt <= 0) OR (nCnt > DL_WMC_N_MAX) THEN
    eErr := DL_WMC_ERR_IN;          // 故障级：nCnt 界外
    bError := TRUE;                 // 故障码配对置位（R101）
    bValid := FALSE;                // 结果不可用
    RETURN;                         // 直接出口 / early exit
END_IF

(* —— 段 3｜单遍累加：非有限元素跳过，守卫计数防失控 —— *)
FOR i := 1 TO nCnt DO
    nGuard := nGuard + 1;           // 守卫递增 / guard increment
    IF nGuard > DL_WMC_GUARD_MAX THEN
        EXIT;                       // 守卫兜底退出（理论不可达）/ guard backstop
    END_IF
    IF (aVals[i] <> aVals[i]) OR (aWeights[i] <> aWeights[i])
       OR ((aVals[i] - aVals[i]) <> (aVals[i] - aVals[i]))
       OR ((aWeights[i] - aWeights[i]) <> (aWeights[i] - aWeights[i])) THEN
        bSkipped := TRUE;           // NaN 自反判 OR Inf 差值自减判：剔除非有限元素
    ELSE
        fNum := fNum + aVals[i] * aWeights[i];   // 分子累加（LREAL 域）/ numerator accumulate
        fWSum := fWSum + aWeights[i];            // 分母累加 / denominator accumulate
    END_IF
END_FOR

(* —— 段 4｜除零防御闸：有效权重和必须 > 阈值 —— *)
IF fWSum <= DL_WMC_TOL THEN
    eErr := DL_WMC_ERR_IN;          // 故障级：权重和为零（防除零拒绝）
    bError := TRUE;                 // 故障码配对置位（R101）
    bValid := FALSE;                // 结果不可用
    RETURN;                         // 直接出口 / early exit
END_IF

(* —— 段 5｜出口 —— *)
FC_DL_WeightedMeanCalc := fNum / fWSum;   // 加权平均（分母已过闸）/ weighted mean
IF bSkipped THEN
    eErr := DL_WMC_INFO_SKIP;       // 信息级：非有限剔除（不置 bError）/ info level
END_IF
bValid := TRUE;                     // 结果可用 / result usable
END_FUNCTION

(* ---- FC_DL_WeightedPercentile.st ---- *)
(*
  ==================================================================
  组件名 Component  : FC_DL_WeightedPercentile
  分类   Category   : DL_MathData
  前缀   Naming     : FC_DL_ ｜ b/n/u/f/t/e/st 类型前缀制（R265）
  复杂度 Complexity  : 中
  版本   Version    : 1.0.1
  功能   Purpose    : 加权百分位数插值（PercentileLReal 升版邻位，权向量参与排序序）。
  来源   Source     : t2-1-lgf-math（LGF Math 百分位族加权变体）
  平台   Platform   : 纯 IEC 61131-3（FOR / 委托 / 四则），三平台通用
  分工声明 Split     : 与 FC_DL_PercentileLReal（等权属主）与 FC_DL_SortIndexLReal
                      （索引排序属主）分工——本件逐级委托后者排序，不重实现
                      排序内核（R140 委托优先，R216 双向互引）。
  依赖     Depends  : FC_DL_SortIndexLReal（DL_MathData 属主，本件委托排序）
  作者   Author     : 道莅代码库 · PLC 编程专家（R61）
  归属 Ownership     : 本件无 TYPE 声明；引用件类型全部 IEC 标准原生。
  ------------------------------------------------------------------
  边界 Boundary     :
                      一 分位 p 钳位 [0,1]：p < 0 钳 0、p > 1 钳 1，置信息级码；
                         p = 0 → 排序首元，p = 1 → 排序末元（两端点向量自证）；
                      二 权向量闸：任一 wᵢ < 0、非有限或 Σw = 0 判故障级拒绝
                         （无权可分即无分位可言）；
                      三 插值除子 (cum_k − cum_{k-1}) ≤ 0 时直接取右元值（禁除零）；
                      四 结果复检兜底同拍置 eErr + bError + bValid 三件套（R258）；
                      五 只读入参数组，不改调用方数据（PercentileLReal 纪律）；
                      六 无状态纯函数：局部量段 1 显式预置（R254）。
  错误码   Codes    :
    16#0001_0639【信息级】计数越域已钳位或分位 p 越域已钳位到 [0,1]
    16#0001_063A【故障级】权向量非法（负权 / 非有限 / Σw = 0），拒绝出值
    16#0001_063B【故障级】结果非有限（复检兜底）
  验收   Acceptance :
    算法已证（脚本）：未跑 ｜ 编译器已证（三平台）：未跑
    V1 值 1/2/3 权 1/1/2、p=0.5 → 目标 2.0 落第 2 位 → 2.0
    V2 p=0 → 首元；p=1 → 末元；p=1.5 → 钳 1 码 0639
    V3 权全零 → 码 063A、bValid=FALSE
    V4 正常 8 样本 → 结果与 v1.0.0 逐位一致（无行为回退，v1.0.1 回归向量）
    V5 委托件返回 TRUE 但内部 bValid=FALSE（构造）→ bSortOk=FALSE（v1.0.1 新增可捕获组合）
  无回退断言 Regression  :
    v1.0.1 仅改委托调用的承接方式（返回值落 _bSortRet、bValid 映射落 _bSortValid，再合取），
    不触碰段 2 / 段 3 / 段 5 / 段 6 的任何判据、钳位与插值公式，故三平台同一输入下
    结果与 v1.0.0 逐位一致（位级相等，非容差相等）。
  修订记录 Revision  :
    2026-11-21  v1.0.0  R61 首版（批 2 · 序号 6）
    2026-11-21  v1.0.1  R62-D5 返修：委托返回值落 _bSortRet、bValid => 落 _bSortValid，再 bSortOk := _bSortRet AND _bSortValid（禁双写同一变量）；头注释补「与 v1.0.0 结果逐位一致」无回退断言说明
  ==================================================================
*)
FUNCTION FC_DL_WeightedPercentile : BOOL
VAR_IN_OUT
    afValues : ARRAY[0..255] OF LREAL; // 数值序列 [工程单位]，只读 / the value series, read only
    afWeights : ARRAY[0..255] OF LREAL; // 权序列 [权]，只读 / the weight series, read only
END_VAR
VAR_INPUT
    nCount : DINT;  // 序列个数 [个]，合法域 1..256 / the count, legal from one to two hundred fifty six
    fP     : LREAL; // 目标分位 [-]，域 [0,1] 钳位 / the target quantile, clamped to the unit domain
END_VAR
VAR_OUTPUT
    fOut   : LREAL; // 加权百分位结果 [工程单位] / the weighted percentile result
    bValid : BOOL;  // 结果可用标志 [-] / the result usable flag
    eErr   : UDINT; // 错误码，0 = 正常 / the error code, zero is ok
    bError : BOOL;  // 错误标志，故障级码置位（R45 配对）/ the error flag
END_VAR
VAR
    aOrd    : ARRAY[0..255] OF DINT; // 排序索引排列（委托输出）/ the sorted permutation from the delegate
    k       : DINT;  // 遍历索引 [下标] / the traversal index
    nUse    : DINT;  // 钳位后的个数 [个] / the clamped count
    fPUse   : LREAL; // 钳位后的分位 [-] / the clamped quantile
    fWsum   : LREAL; // 权和 [权] / the weight sum
    fTarget : LREAL; // 目标累积权 [权] / the target cumulative weight
    fCum    : LREAL; // 当前累积权 [权] / the current cumulative weight
    fCumPrv : LREAL; // 前一位置累积权 [权] / the previous cumulative weight
    fVL     : LREAL; // 插值左元值 [工程单位] / the left interpolation value
    fVR     : LREAL; // 插值右元值 [工程单位] / the right interpolation value
    fFrac   : LREAL; // 插值分数 [-] / the interpolation fraction
    nHit    : DINT;  // 命中位置 [下标] / the hit position
    bFound  : BOOL;  // 命中标记 [-] / the hit flag
    bSortOk : BOOL;  // 委托排序可用位（返回值与 bValid 合取）/ the delegate sort usable bit, the conjunction
    _bSortRet : BOOL; // 委托函数返回值承接变量（独立承接，禁双写，R62-D5）/ the delegate return value holder, never double written
    _bSortValid : BOOL; // 委托 bValid 输出承接变量（独立承接，禁双写）/ the delegate valid output holder, never double written
    bSortEr : BOOL;  // 委托排序故障位 [-] / the delegate sort fault bit
    uSortEr : UDINT; // 委托排序错误码 [码] / the delegate error code
    bClamp  : BOOL;  // 钳位发生标记 [-] / the clamp happened flag
END_VAR
VAR CONSTANT
    DL_WPC_NMAX : DINT := 256; // 序列容量上界 [个]，与数组容量一致 / the capacity aligned with the array
END_VAR

// 段 1｜返回值与错误状态预置安全值 + 局部量显式预置（R45 / R254）/ segment 1, the preset
FC_DL_WeightedPercentile := FALSE; // 返回值预置假 / preset the return false
fOut := 0.0; // 结果预置零 / preset the result zero
bValid := FALSE; // 有效标志预置假 / preset the validity false
eErr := 16#0000_0000; // 错误码预置正常 / preset the code to ok
bError := FALSE; // 错误标志预置假 / preset the error flag false
nUse := 0; // 个数预置零 / preset the count zero
fPUse := 0.0; // 分位预置零 / preset the quantile zero
fWsum := 0.0; // 权和预置零 / preset the weight sum zero
fTarget := 0.0; // 目标累积权预置零 / preset the target zero
fCum := 0.0; // 累积权预置零 / preset the cumulative zero
fCumPrv := 0.0; // 前位累积权预置零 / preset the previous zero
fVL := 0.0; // 左元值预置零 / preset the left value zero
fVR := 0.0; // 右元值预置零 / preset the right value zero
fFrac := 0.0; // 分数预置零 / preset the fraction zero
nHit := 0; // 命中位置预置零 / preset the hit zero
bFound := FALSE; // 命中标记预置假 / preset the hit flag false
bSortOk := FALSE; // 委托成功位预置假 / preset the delegate bit false
_bSortRet := FALSE; // 委托返回值承接量预置假 / preset the return holder false
_bSortValid := FALSE; // 委托可用位承接量预置假 / preset the valid holder false
bSortEr := FALSE; // 委托故障位预置假 / preset the delegate fault bit false
uSortEr := 16#0000_0000; // 委托码预置零 / preset the delegate code zero
bClamp := FALSE; // 钳位标记预置假 / preset the clamp flag false
FOR k := 0 TO 255 DO // 排列数组预置恒等 / preset the permutation array
    aOrd[k] := k; // 恒等索引 / the identity index
END_FOR

// 段 2｜计数与分位域闸（钳位显式，边界一）/ segment 2, the count and quantile gates
IF nCount < 1 THEN // 空序列无分位 / an empty series has no percentile
    eErr := 16#0001_0639; // 信息级：计数越域已钳位（信息级不置 bError）/ informational, the count clamped
    RETURN; // 早退：fOut 保持零、bValid 保持假 / early return
END_IF
nUse := nCount; // 域内接管 / take the count
IF nUse > DL_WPC_NMAX THEN // 超容量 / above the capacity
    nUse := DL_WPC_NMAX; // 钳到容量 / clamp to the capacity
    bClamp := TRUE; // 置钳位标记 / raise the clamp flag
END_IF
fPUse := fP; // 分位接管 / take the quantile
IF fPUse < 0.0 THEN // 低于下界 / below the floor
    fPUse := 0.0; // 钳到零 / clamp to zero
    bClamp := TRUE; // 置钳位标记 / raise the clamp flag
END_IF
IF fPUse > 1.0 THEN // 高于上界 / above the ceiling
    fPUse := 1.0; // 钳到一 / clamp to one
    bClamp := TRUE; // 置钳位标记 / raise the clamp flag
END_IF
IF (fPUse <> fPUse) OR ((fPUse - fPUse) <> (fPUse - fPUse)) THEN // 分位非有限（NaN 钳位序闸兜不住，逐个点名，R272）/ a non finite quantile
    eErr := 16#0001_063A; // 故障级：入参非法归权向量闸同码口径（判据集合内非法）/ fault grade, an illegal input
    bError := TRUE; // 置错误标志（R45 配对）/ raise the error flag
    RETURN; // 早退 / early return
END_IF
IF bClamp THEN // 钳位发生置信息级 / the clamp raises the informational code
    eErr := 16#0001_0639; // 信息级：计数或分位越域已钳位 / informational, clamped
END_IF

// 段 3｜权向量闸：逐元素负权 / 非有限点名 + Σw 判（边界二，R272）/ segment 3, the weight gate
FOR k := 0 TO nUse - 1 DO // 有界遍历 / the bounded traversal
    IF (afWeights[k] < 0.0)
    OR (afWeights[k] <> afWeights[k])
    OR ((afWeights[k] - afWeights[k]) <> (afWeights[k] - afWeights[k])) THEN // 负权或非有限 / a negative or non finite weight
        eErr := 16#0001_063A; // 故障级：权向量非法 / fault grade, an illegal weight vector
        bError := TRUE; // 置错误标志（R45 配对）/ raise the error flag
        RETURN; // 早退 / early return
    END_IF
    fWsum := fWsum + afWeights[k]; // 权和累加 / accumulate the weight sum
END_FOR
IF fWsum <= 0.0 THEN // 权和为零（权和已证非负，本判覆盖恰零）/ a zero weight sum
    eErr := 16#0001_063A; // 故障级：权向量和为零 / fault grade, the zero weight sum
    bError := TRUE; // 置错误标志（R45 配对）/ raise the error flag
    RETURN; // 早退 / early return
END_IF

// 段 4｜委托稳定排序（R140 委托优先；返回值与 bValid 分承，禁双写，R62-D5）/ segment 4, the delegated stable sort with two separate holders
_bSortRet := FC_DL_SortIndexLReal(afValues := afValues, nCount := nUse, aIdx => aOrd, bValid => _bSortValid, eErr => uSortEr, bError => bSortEr); // 委托索引排序：返回值落 _bSortRet、可用位映射落 _bSortValid / delegate the index sort with two distinct holders
bSortOk := _bSortRet AND _bSortValid; // 返回值与可用位各自承接后合取（IEC 未规定返回值与输出映射的求值次序）/ conjoin the return value and the valid flag, since IEC leaves their evaluation order unspecified
IF (NOT bSortOk) OR bSortEr THEN // 委托失败（含其非有限故障码回传）/ the delegate failed
    eErr := uSortEr; // 委托码回传（码随属主，R66）/ replay the delegate code
    bError := bSortEr; // 委托故障位回传 / replay the delegate fault bit
    RETURN; // 早退 / early return
END_IF

// 段 5｜加权累积定位与邻位插值（边界一三）/ segment 5, the weighted location and the neighbour interpolation
fTarget := fPUse * fWsum; // 目标累积权（p=0 取首元、p=1 取末元，两端点自证）/ the target cumulative weight
fCum := 0.0; // 累积权清零 / reset the cumulative
FOR k := 0 TO nUse - 1 DO // 按排序序累积（命中后余轮守卫跳过，禁改循环变量）/ accumulate in the sorted order, the rounds after the hit are guarded out
    IF NOT bFound THEN // 未命中才继续累积 / accumulate only before the hit
        fCumPrv := fCum; // 前位累积权快照 / snapshot the previous cumulative
        fCum := fCum + afWeights[aOrd[k]]; // 累进当前权 / add the current weight
        IF fCum >= fTarget THEN // 越过目标即命中（p=0 时首位置即命中）/ the target crossed
            nHit := k; // 记录命中位置 / register the hit position
            bFound := TRUE; // 置命中标记 / raise the hit flag
        END_IF
    END_IF
END_FOR
IF NOT bFound THEN // 全遍历未越过（浮点和误差兜底）：取末元 / the fallback to the last element
    nHit := nUse - 1; // 命中末位置 / the last position
END_IF
fVR := afValues[aOrd[nHit]]; // 右元值 = 命中位值 / the right value is the hit value
IF nHit = 0 THEN // 命中首位：无左邻（p=0 端点）/ the first position, no left neighbour
    fOut := fVR; // 直接取右元 / take the right value directly
ELSE // 邻位插值 / the neighbour interpolation
    fVL := afValues[aOrd[nHit - 1]]; // 左元值 / the left value
    IF (fCum - fCumPrv) > 0.0 THEN // 插值除子已证 > 0（边界三）/ the proven positive divisor
        fFrac := (fTarget - fCumPrv) / (fCum - fCumPrv); // 插值分数 / the interpolation fraction
        IF fFrac < 0.0 THEN // 分数越下界（浮点和误差兜底钳位）/ the fraction below the floor
            fFrac := 0.0; // 钳到零（取左元）/ clamp to zero
        END_IF
        IF fFrac > 1.0 THEN // 分数越上界 / the fraction above the ceiling
            fFrac := 1.0; // 钳到一（取右元）/ clamp to one
        END_IF
        fOut := fVL + (fVR - fVL) * fFrac; // 线性插值出结果 / the linear interpolation
    ELSE // 除子非正（零权相邻）：直接取右元（禁除零，边界三）/ a non positive divisor, take the right value
        fOut := fVR; // 直接取右元 / take the right value directly
    END_IF
END_IF

// 段 6｜结果复检兜底（非有限同拍三件套，边界四）/ segment 6, the result recheck
IF (fOut <> fOut) OR ((fOut - fOut) <> (fOut - fOut)) THEN // 结果非有限 / the result is not finite
    fOut := 0.0; // 兜底安全值 / the bottom line safe value
    eErr := 16#0001_063B; // 故障级：结果非有限 / fault grade, the non finite result
    bError := TRUE; // 置错误标志（R45 配对）/ raise the error flag
    bValid := FALSE; // 结果不可用 / the result void
    RETURN; // 早退 / early return
END_IF
bValid := TRUE; // 结果可用 / the result is usable
FC_DL_WeightedPercentile := TRUE; // 返回成功 / return success
END_FUNCTION

(* ---- FC_DL_WeirFlowCalc.st ---- *)
(*
  道莅工业代码库 | DL_MathData | FC_DL_WeirFlowCalc
  版本: 1.0.0 | 日期: 2026-11-23 | 轮次: R75
  开源溯源: self-cleanroom（无外部来源；薄壁堰/宽顶堰过流公式为水力学公开公式，零代码行复制）
  功能: 堰流过流量计算——薄壁堰 Q = (2/3)·Cd·b·√(2g)·hu^1.5 与宽顶堰
        Q = Mb·b·√(2g)·hu^1.5，含淹没流判别（hd/hu > 阈值）与淹没折减因子。
  兼容性: CODESYS 3.5 / TwinCAT 3 / 汇川 InoProShop；仅依赖标准 SQRT/ABS，零厂商私有库
  接口: 输入堰上水头/堰下（下游）水头/堰宽/堰型/两系数/淹没判别比；函数返回值
        = 过流量 [m3/s]（非法入参返回 0.0），输出 bSubmerged/bValid/eErr。
        纯函数：无内部状态，每拍独立全量重算。
  码表: 16#0001_03FF 故障级：入参域非法（水头/宽度/系数越域或非有限）→ bValid=FALSE
        码段说明：0001 段故障子带 03xx，03FF 槽经全库实扫空闲。
  边界: ① 域闸：hu > 0、b > 0、Cd > 0、Mb > 0、0 < 淹没比 < 1，全部入参 NaN 自反判；
        ② 淹没判别 hd/hu 除法前由 hu > 0 域闸保证；
        ③ 淹没折减因子 √(1 - r^1.5) 底数用 MAX(0, ·) 钳非负，杜绝负数开方；
        ④ hu^1.5 以 hu·√hu 实现（同幂等价，免 EXPT 泛型疑义）；
        ⑤ 全部输出在所有路径（含提前返回）赋值；⑥ 零全局耦合。
  邻件比对: OrificeFlowCalc（孔口流 vs 堰流，公式域不同）。
  修订历史: 2026-11-23 v1.0.0 R75 首版（复杂件批 B2 · C06）
*)

FUNCTION FC_DL_WeirFlowCalc : REAL
VAR_INPUT
    fHeadUp     : REAL := 0.0;    // 堰上水头（高于堰顶），域 > 0 [m] | Upstream head above crest
    fHeadDown   : REAL := 0.0;    // 堰下（下游）水头（高于堰顶）[m] | Downstream head above crest
    fWidth      : REAL := 1.0;    // 堰宽（垂直流向有效宽度），域 > 0 [m] | Weir crest width
    bBroadCrest : BOOL := FALSE;  // 堰型选择：TRUE=宽顶堰，FALSE=薄壁堰 [-] | TRUE = broad-crested, FALSE = thin-plate
    fCd         : REAL := 0.611;  // 薄壁堰流量系数，域 > 0 [-] | Thin-plate discharge coefficient
    fMb         : REAL := 0.36;   // 宽顶堰流量系数，域 > 0 [-] | Broad-crested discharge coefficient
    fSubmRatio  : REAL := 0.75;   // 淹没判别比阈值，域 (0, 1) [-] | Submergence ratio threshold
END_VAR
VAR_OUTPUT
    bSubmerged : BOOL;            // 本拍淹没流判别结果 [-] | Submerged flow judgement
    bValid     : BOOL;            // 本次计算有效 [-] | Computation valid
    eErr       : UDINT;           // 错误码，0 = 无错 | Error code, 0 = none
END_VAR
VAR
    fHu15    : REAL;              // 堰上水头 1.5 次幂 hu^1.5 [m^1.5] | Upstream head to power 1.5
    fRatio   : REAL;              // 淹没比 hd/hu [-] | Submergence ratio
    fRatio15 : REAL;              // 淹没比 1.5 次幂 r^1.5 [-] | Ratio to power 1.5
    fFactor  : REAL;              // 淹没折减因子 [-] | Submergence reduction factor
    fCoef    : REAL;              // 按堰型选定的合成系数 [-] | Combined coefficient by weir type
    fQ       : REAL;              // 过流量暂存 [m3/s] | Flow staging
    bInOk    : BOOL;              // 入参域合法当拍量 [-] | Input domain legal this call
END_VAR
VAR CONSTANT
    DL_WFC_G2   : REAL := 19.62;      // 重力加速度二倍 2g [m/s2] | Twice gravity
    DL_WFC_EPS  : REAL := 1.0E-6;     // 判零容差（水头/宽度近零判据） | Zero threshold tolerance
    DL_WFC_ERR  : UDINT := 16#0001_03FF;  // 入参域非法码 | Illegal input domain code
END_VAR

(* —— 段 0：输出缺省全赋值（全路径覆盖） —— *)
bSubmerged := FALSE;              // 淹没判别预置 FALSE / Submerged preset FALSE
bValid := FALSE;                  // 有效标志预置 FALSE / Valid preset FALSE
eErr := 0;                        // 错误码缺省 / Error default
fQ := 0.0;                        // 流量暂存清零（防御） / Flow staging cleared
FC_DL_WeirFlowCalc := 0.0;        // 返回值缺省零（非法路径出口） / Return default zero

(* —— 段 1：入参域闸（NaN 自反判 + 域上下界） —— *)
bInOk := (fHeadUp > DL_WFC_EPS) AND (fWidth > DL_WFC_EPS)
      AND (fCd > 0.0) AND (fMb > 0.0)
      AND (fSubmRatio > 0.0) AND (fSubmRatio < 1.0)
      AND (fHeadUp = fHeadUp) AND (fHeadDown = fHeadDown)
      AND (fWidth = fWidth) AND (fCd = fCd) AND (fMb = fMb) AND (fSubmRatio = fSubmRatio);
IF NOT bInOk THEN
    eErr := DL_WFC_ERR;           // 域非法码 / Domain illegal code
    RETURN;                       // 提前返回：输出已全赋值 / Early return, outputs assigned
END_IF

(* —— 段 2：淹没判别（除法分母 hu > EPS 已由域闸证明） —— *)
fRatio := fHeadDown / fHeadUp;    // 淹没比 hd/hu / Submergence ratio
bSubmerged := fRatio > fSubmRatio;  // 淹没判别 / Submerged judgement
IF fRatio < 0.0 THEN
    fRatio := 0.0;                // 负下游水头（低于堰顶）钳零 / Negative downstream head clamped
END_IF

(* —— 段 3：过流量主式（按堰型选系数） —— *)
fHu15 := fHeadUp * SQRT(fHeadUp); // hu^1.5 = hu·√hu / Head to power 1.5
IF bBroadCrest THEN
    fCoef := fMb;                 // 宽顶堰系数 / Broad-crested coefficient
ELSE
    fCoef := (2.0 / 3.0) * fCd;   // 薄壁堰系数 (2/3)·Cd / Thin-plate coefficient
END_IF
fQ := fCoef * fWidth * SQRT(DL_WFC_G2) * fHu15;   // 自由出流过流量 [m3/s] / Free flow discharge

(* —— 段 4：淹没折减（因子底数钳非负，杜绝负数开方） —— *)
IF bSubmerged THEN
    fRatio15 := fRatio * SQRT(fRatio);                  // r^1.5 = r·√r（r ≥ 0 已钳）/ Ratio to power 1.5
    fFactor := SQRT(MAX(0.0, 1.0 - fRatio15));          // 折减因子 ∈ [0, 1] / Reduction factor clamped non-negative
    fQ := fQ * fFactor;                                 // 淹没过流量 [m3/s] / Submerged discharge
END_IF

(* —— 段 5：出口赋值 —— *)
FC_DL_WeirFlowCalc := fQ;         // 返回过流量 [m3/s] / Return discharge
bValid := TRUE;                   // 计算有效 / Valid

END_FUNCTION

(* ---- FC_DL_WetBulbCalc.st ---- *)
(*
  Name        : FC_DL_WetBulbCalc
  Category    : DL_MathData
  Version     : 1.0.0
  Purpose     : 干球温度/相对湿度的湿球温度迭代估算：以 Magnus 饱和水汽压式构造热力学方程，牛顿迭代求根（焓湿图原子补口）；/ Wet-bulb temperature estimation from dry-bulb temperature and relative humidity: Magnus saturation-vapour formulation solved by Newton iteration
  溯源        : 借 t1-2-oscat-building 的分类/参数域组织，clean-room 实现
  Boundary    : ① 入口有限性闸：任一输入 NaN（x = x 自反）或 Inf（(x-x) = (x-x) 差判）→ bValid = FALSE，返回 0.0（哨兵零点，不饱和、不外推）；
                ② 输入域钳位：干球温度钳 -40..80 °C、相对湿度钳 1..100 %、气压钳 300..1100 hPa，钳位是各自中间量的最后一次写；
                ③ 牛顿迭代：上限 20 次，步长收敛阈 DL_WBC_EPS；迭代发散（导数近零）即刻退出并置 bValid = FALSE；
                ④ 除零前置：迭代导数 |des + gamma| < eps 时不除（发散路径）；湿度换算除子为常量 100.0；
                ⑤ 返回值 = 湿球温度 [°C]，bValid = FALSE 时不得使用返回值（上层契约）。
*)
FUNCTION FC_DL_WetBulbCalc : REAL
VAR_INPUT
    fTempDry  : REAL;                        (* 干球温度 [°C] / Dry-bulb temperature *)
    fRelHum   : REAL;                        (* 相对湿度，域 1..100（越域钳位）[%] / Relative humidity, clamped *)
    fPressure : REAL := 1013.25;             (* 大气压，域 300..1100（越域钳位）[hPa] / Atmospheric pressure, clamped *)
END_VAR
VAR_OUTPUT
    bValid    : BOOL;                        (* 结果有效标志（FALSE 时返回值为哨兵零点）[-] / Result validity flag *)
END_VAR
VAR
    _fT       : REAL;                        (* 钳位后干球温度中间量 [°C] / Clamped dry-bulb temperature *)
    _fRh      : REAL;                        (* 钳位后相对湿度中间量 [%] / Clamped relative humidity *)
    _fP       : REAL;                        (* 钳位后气压中间量 [hPa] / Clamped pressure *)
    _fEs      : REAL;                        (* 干球温度饱和水汽压 [Pa] / Saturation vapour pressure at dry bulb *)
    _fE       : REAL;                        (* 实际水汽压 [Pa] / Actual vapour pressure *)
    _fGamma   : REAL;                        (* 湿计常数 gamma = 0.00066 × P [Pa/°C 口径见实现] / Psychrometric constant *)
    _fTw      : REAL;                        (* 湿球温度迭代变量 [°C] / Wet-bulb iterate *)
    _fEsW     : REAL;                        (* 湿球温度饱和水汽压 [Pa] / Saturation vapour pressure at wet bulb *)
    _fDesW    : REAL;                        (* 饱和水汽压对湿球温度导数 [Pa/°C] / Derivative of es at wet bulb *)
    _fFv      : REAL;                        (* 方程残差 f(Tw) [Pa] / Equation residual *)
    _fDv      : REAL;                        (* 方程导数 f'(Tw) [Pa/°C] / Equation derivative *)
    _fStep    : REAL;                        (* 牛顿步长（绝对值判敛）[°C] / Newton step magnitude *)
    _nIt      : INT;                         (* 迭代计数 [次] / Iteration counter *)
    _bOk      : BOOL;                        (* 求解成功内部量 / Solve-success internal *)
END_VAR
VAR CONSTANT
    DL_WBC_EPS   : REAL := 1.0E-4;           (* 迭代收敛阈值 [°C] / Convergence threshold *)
    DL_WBC_ITMAX : INT  := 20;               (* 牛顿迭代上限 [次] / Newton iteration cap *)
    DL_WBC_A     : REAL := 17.625;           (* Magnus 系数 a [-] / Magnus coefficient a *)
    DL_WBC_B     : REAL := 243.04;           (* Magnus 系数 b [°C] / Magnus coefficient b *)
    DL_WBC_ES0   : REAL := 610.94;           (* Magnus 基准饱和水汽压 [Pa] / Magnus base saturation pressure *)
    DL_WBC_HUND  : REAL := 100.0;            (* 湿度百分数换算常量（常量除子）[-] / Percent scale constant *)
    DL_WBC_TMIN  : REAL := -40.0;            (* 干球温度钳位下限 [°C] / Dry-bulb clamp floor *)
    DL_WBC_TMAX  : REAL := 80.0;             (* 干球温度钳位上限 [°C] / Dry-bulb clamp ceiling *)
    DL_WBC_PMIN  : REAL := 300.0;            (* 气压钳位下限 [hPa] / Pressure clamp floor *)
    DL_WBC_PMAX  : REAL := 1100.0;           (* 气压钳位上限 [hPa] / Pressure clamp ceiling *)
END_VAR

(* —— 段 0：入口有限性闸（NaN 自反 + Inf 差判，三输入逐项） —— *)
bValid := TRUE;                                                                (* 有效标志预置（任一闸命中即翻 FALSE） / Validity preset *)
IF NOT ((fTempDry = fTempDry) AND ((fTempDry - fTempDry) = (fTempDry - fTempDry))) THEN
    bValid := FALSE;                                                           (* 干球温度非有限 / Dry bulb non-finite *)
END_IF
IF NOT ((fRelHum = fRelHum) AND ((fRelHum - fRelHum) = (fRelHum - fRelHum))) THEN
    bValid := FALSE;                                                           (* 相对湿度非有限 / Humidity non-finite *)
END_IF
IF NOT ((fPressure = fPressure) AND ((fPressure - fPressure) = (fPressure - fPressure))) THEN
    bValid := FALSE;                                                           (* 气压非有限 / Pressure non-finite *)
END_IF

(* —— 段 1：无效输入早退（返回哨兵零点，不饱和、不外推） —— *)
IF NOT bValid THEN
    FC_DL_WetBulbCalc := 0.0;                                                  (* 哨兵零点返回 / Sentinel zero return *)
    RETURN;
END_IF

(* —— 段 2：输入域钳位（各自中间量最后一次写，钳位不被覆盖） —— *)
_fT := fTempDry;                                                               (* 干球温度装载 / Load dry bulb *)
IF _fT < DL_WBC_TMIN THEN
    _fT := DL_WBC_TMIN;                                                        (* 下限钳位 / Lower clamp *)
END_IF
IF _fT > DL_WBC_TMAX THEN
    _fT := DL_WBC_TMAX;                                                        (* 上限钳位 / Upper clamp *)
END_IF
_fRh := fRelHum;                                                               (* 相对湿度装载 / Load humidity *)
IF _fRh < 1.0 THEN
    _fRh := 1.0;                                                               (* 湿度下限钳 1（防 0 湿度发散） / Humidity lower clamp *)
END_IF
IF _fRh > DL_WBC_HUND THEN
    _fRh := DL_WBC_HUND;                                                       (* 湿度上限钳 100 / Humidity upper clamp *)
END_IF
_fP := fPressure;                                                              (* 气压装载 / Load pressure *)
IF _fP < DL_WBC_PMIN THEN
    _fP := DL_WBC_PMIN;                                                        (* 气压下限钳位 / Pressure lower clamp *)
END_IF
IF _fP > DL_WBC_PMAX THEN
    _fP := DL_WBC_PMAX;                                                        (* 气压上限钳位 / Pressure upper clamp *)
END_IF

(* —— 段 3：热力学方程构造（Magnus + 湿计方程） —— *)
_fEs := DL_WBC_ES0 * EXP(DL_WBC_A * _fT / (_fT + DL_WBC_B));                   (* 干球温度饱和水汽压（除子 _fT+243.04 恒 > 0，域钳位保证）[Pa] / es at dry bulb *)
_fE := _fRh / DL_WBC_HUND * _fEs;                                             (* 实际水汽压（除子为常量）[Pa] / Actual vapour pressure *)
_fGamma := 0.00066 * _fP;                                                     (* 湿计常数（无除法）[hPa/°C] / Psychrometric constant *)

(* —— 段 4：牛顿迭代求湿球温度（发散与不收敛均落 bValid = FALSE，安全侧） —— *)
_fTw := _fT;                                                                   (* 迭代初值取干球温度（物理上界） / Init at dry bulb *)
_bOk := FALSE;                                                                 (* 求解成功内部量预清 / Success preset *)
_nIt := 0;                                                                     (* 迭代计数清零 / Counter clear *)
WHILE _nIt < DL_WBC_ITMAX DO
    _fEsW := DL_WBC_ES0 * EXP(DL_WBC_A * _fTw / (_fTw + DL_WBC_B));            (* 湿球温度饱和水汽压 [Pa] / es at wet bulb *)
    _fDesW := _fEsW * DL_WBC_A * DL_WBC_B / ((_fTw + DL_WBC_B) * (_fTw + DL_WBC_B));   (* Magnus 导数（除子平方项恒 > 0）[Pa/°C] / Derivative of es *)
    _fFv := _fEsW - _fGamma * (_fT - _fTw) - _fE;                              (* 残差 f(Tw) = es(Tw) - gamma·(T - Tw) - e [Pa] / Residual *)
    _fDv := _fDesW + _fGamma;                                                  (* 导数 f'(Tw)（湿计项恒正）[Pa/°C] / Derivative *)
    IF ABS(_fDv) < DL_WBC_EPS THEN
        _bOk := FALSE;                                                         (* 导数近零：发散退出（除零前置，边界③） / Diverged on near-zero derivative *)
        EXIT;
    END_IF
    _fStep := _fFv / _fDv;                                                     (* 牛顿步长（除子已过闸）[°C] / Newton step *)
    _fTw := _fTw - _fStep;                                                     (* 迭代递进 / Iterate advance *)
    IF _fTw > _fT THEN
        _fTw := _fT;                                                           (* 湿球不超干球（物理上界钳位） / Wet bulb <= dry bulb *)
    END_IF
    IF _fTw < _fT - 60.0 THEN
        _fTw := _fT - 60.0;                                                    (* 湿球下界钳位（防迭代飞逸） / Wet bulb floor *)
    END_IF
    IF ABS(_fStep) < DL_WBC_EPS THEN
        _bOk := TRUE;                                                          (* 步长收敛：求解成功 / Converged *)
        EXIT;
    END_IF
    _nIt := _nIt + 1;                                                          (* 迭代计数递进 / Counter advance *)
END_WHILE

(* —— 段 5：出口（bValid 由收敛结果定，返回湿球温度） —— *)
bValid := _bOk;                                                                (* 有效标志 = 收敛成功 / Validity = converged *)
IF bValid THEN
    FC_DL_WetBulbCalc := _fTw;                                                 (* 湿球温度返回 [°C] / Wet-bulb return *)
ELSE
    FC_DL_WetBulbCalc := 0.0;                                                  (* 未收敛返回哨兵零点（安全侧契约） / Sentinel zero on divergence *)
END_IF
END_FUNCTION

(* ---- FC_DL_WordFromBytes.st ---- *)
(*==============================================================================
 * 组件名称 (Component)  : FC_DL_WordFromBytes
 * 所属子库 (Sublibrary) : DL_MathData
 * 当前版本 (Version)    : 1.0.0
 * 兼容性   (Platform)   : CODESYS 3.5 / TwinCAT 3 / 汇川 InoProShop / Machine Expert
 *                         仅依赖 Standard.library（SHL / AND / OR / 类型转换），零厂商方言
 * 来源标签 (Source)     : t2-1-lgf-converter（字节序组装族，clean-room 编写）
 * 功能描述 (Function)   : BYTE 数组按字节序组装为 WORD / DWORD。返回值以 DWORD 承载：
 *                         nTargetLen = 2 时结果在低 16 位（高 16 位恒零），
 *                         nTargetLen = 4 时为完整 32 位结果。
 *                         四序语义（E_DL_ByteOrder，WORD 目标下三序退化披露）：
 *                           eAbcd：字节 i 落槽位 i（槽 0 = 最高字节，大端直排）
 *                           eDcba：字节 i 落槽位 (nTargetLen-1-i)（全反序）
 *                           eBadc：字节 i 落槽位 (i XOR 1)（寄存器内两两互换）
 *                           eCdab：DWORD 下字节 i 落槽位 (i XOR 2)（高低字互换）；
 *                                  WORD 下退化为字节反序（单字容器内高低字互换
 *                                  不可区分，验收向量 16#1234 即按此口径）。
 *                         组装字节数不足按高段补零并置信息级；映射为对合（ involutive），
 *                         与 FC_DL_WordToBytes 同序构成 round-trip 双向对。
 * 归属声明 (Ownership)  : E_DL_ByteOrder 归属 DL_MathData\FC_DL_SwapBytes32.st，
 *                         本件只引用不重声明（FB51-7）。
 * 边界与语义披露 (Boundary disclosure) :
 *   1) 指针 NIL 或字节数 <= 0：结构性早退，返回零值 + bValid FALSE（零写入语义），
 *      不触碰调用方内存。
 *   2) 组装字节数大于目标长度：多余低位字节忽略（不计码——调用方传入 nCount
 *      本身即可观测该事实，R90 反证成立不加码）。
 *   3) 移位量上界 (nTargetLen-1-slot)*8 结构性 <= 24 < 32（DWORD 位宽），禁 MOD
 *      归一的不变量由本披露承担（R48 口径：非裸变量超宽移位）。
 *   4) 验收向量：CDAB 序 {16#34, 16#12} -> 16#0000_1234；ABCD {16#12,16#34,16#56,16#78}
 *      -> 16#1234_5678；长度 1 组装 WORD -> 16#0000_1200 高段补零 + 信息级。
 * 故障码表 (Error codes) :
 *   16#0001_03F3 [故障级] 字节指针 NIL 或 nCount <= 0，返回零 + bValid FALSE
 *                 反证：零返回值与「源字节全零」的正常结果组合相同，bValid
 *                 只表达有效性，故障成因必须由码位承载。
 *   16#0001_03F4 [故障级] 字节序枚举越界（非 0..3），回退默认大端 eAbcd 继续服务
 *                 （对齐 Crc8 非法变体先例：先落默认行为再置码）
 *                 反证：eAbcd 回退结果与显式填 eAbcd 输出组合相同，码位承载
 *                 「组态有误」事实。
 *   16#0001_04B8 [信息级] 源字节数不足目标长度，高段槽位补零
 *                 反证：补零结果与「源字节高段本来就是零」组合相同，无码不可区分。
 *   16#0001_04B9 [信息级] nTargetLen 非 2/4，回退默认 WORD（2 字节）继续服务
 *                 反证：回退结果与显式填 2 相同，码位承载组态有误事实。
 * 码位总账 (Code ledger) : 16#0001_03F3 / 03F4 用 ｜ 16#0001_04B8 / 04B9 用
 * 依赖     (Depends)    : TYPE E_DL_ByteOrder（属主 FC_DL_SwapBytes32.st，只引用）
 * 红线自检 (Redline)    : R1 ✓ 零全局变量与 VAR_EXTERNAL ｜ R2 ✓ 零 %I/%Q 物理地址
 *                         R3 ✓ 纯 IEC 61131-3（指针判空 + 标准移位/转换）
 *                         R4 ✓ 指针 NIL 闸 / 计数域闸 / 枚举域闸 / 全分支码位配对
 *                         R5 ✓ 全变量中英双语同行注释 ｜ R6 N/A（纯函数，无状态机）
 *                         R7 N/A（无定时器 / 边沿实例）
 * 修订历史 (Revision)   :
 *   2026-11-22  v1.0.0  首版入库（R68 构建轮 · 批 1 · 目标 4）
 *============================================================================*)
FUNCTION FC_DL_WordFromBytes : DWORD
VAR_INPUT
    pBytes     : POINTER TO BYTE;   // 源字节数组首指针，NIL = 无效 / Source byte pointer, NIL invalid
    nCount     : INT;               // 源字节数 [个]，<= 0 无效 / Source byte count, <= 0 invalid
    eOrder     : E_DL_ByteOrder;    // 字节序选择（属主 FC_DL_SwapBytes32.st）/ Byte order selector
    nTargetLen : INT := 2;          // 目标长度 [字节]，2 = WORD，4 = DWORD / Target length in bytes
END_VAR
VAR_OUTPUT
    bValid   : BOOL;    // 本拍组装有效 / Assembly valid this call
    bError   : BOOL;    // 故障标志（0305 / 0306 置位，R45 配对）/ Fault flag, set on 0305 and 0306
    uInfoId  : UDINT;   // 故障码，0 = 无故障（纯函数每拍重算）/ Error code, recomputed per call
END_VAR
VAR
    uAcc     : DWORD;   // 组装累加器 / Assembly accumulator
    nUse     : INT;     // 实际参与组装的字节数 [个] / Bytes actually assembled
    nSlot    : INT;     // 当前字节映射到的槽位 [0..3] / Slot the current byte maps to
    nShift   : DINT;    // 当前槽位移位量 [bit]，结构性 <= 24（ANY_INT 口径）/ Slot shift, structurally <= 24
    uB       : BYTE;    // 当前源字节 / Current source byte
    nLenUse  : INT;     // 钳位后的目标长度 [字节] / Clamped target length
    bOrderOk : BOOL;    // 字节序枚举合法性 / Byte order validity
    i        : INT;     // 遍历索引 / Loop index
END_VAR
VAR CONSTANT
    DL_WFB_LEN_MIN : INT := 2;    // 目标长度下限 [字节]（WORD）/ Target length floor, WORD
    DL_WFB_LEN_MAX : INT := 4;    // 目标长度上限 [字节]（DWORD）/ Target length ceiling, DWORD
END_VAR

(*------------------------------------------------------------------------------
 * 段 1｜安全预置（P-01 范式）：任何异常路径返回零 + bValid FALSE，绝不返回残值
 *      Safe preset: every exceptional path returns zero with bValid FALSE
 *-----------------------------------------------------------------------------*)
FC_DL_WordFromBytes := 16#0000_0000;
bValid  := FALSE;
bError  := FALSE;
uInfoId := 16#0000_0000;

(*------------------------------------------------------------------------------
 * 段 2｜域闸（R151 全枚举：指针 + 计数 + 目标长度 + 枚举四闸，结构性 IF/ELSE 不用 RETURN）
 *      Domain gates: pointer, count, target length and enum, full IF/ELSE coverage
 *-----------------------------------------------------------------------------*)
IF (pBytes = 0) OR (nCount <= 0) THEN
    uInfoId := 16#0001_03F3;    // 故障级：指针 NIL 或计数非法 / Fault: NIL pointer or bad count
    bError  := TRUE;            // R45 配对：故障码同行置位 / Paired with the fault code
    RETURN;                     // 结构性早退：输出已全预置，零写入语义成立（规格明示豁免）
END_IF

IF (nTargetLen < DL_WFB_LEN_MIN) OR (nTargetLen > DL_WFB_LEN_MAX) THEN
    nLenUse := DL_WFB_LEN_MIN;  // 二级回退：钳回默认 WORD（R117 两级参数回退）
    uInfoId := 16#0001_04B9;    // 信息级：目标长度非法回默认 / Info: length defaulted
ELSE
    nLenUse := nTargetLen;      // 合法直通 / Valid pass-through
END_IF

bOrderOk := (eOrder = E_DL_ByteOrder.eAbcd) OR (eOrder = E_DL_ByteOrder.eDcba)
            OR (eOrder = E_DL_ByteOrder.eBadc) OR (eOrder = E_DL_ByteOrder.eCdab);
IF NOT bOrderOk THEN
    uInfoId := 16#0001_03F4;    // 故障级：字节序越界回默认大端（0142 风格先例口径）/ Fault: order defaulted
    bError  := TRUE;            // R45 配对 / Paired with the fault code
END_IF

(*------------------------------------------------------------------------------
 * 段 3｜组装主体（边界 B1/B3）：映射 -> 取字节 -> 升位 -> 移位 -> 或合
 *      Assembly body: map, fetch, widen, shift, OR-accumulate
 *      nUse 不足 nLenUse 时高位槽不落值 = 高段补零（信息级 0407）
 *-----------------------------------------------------------------------------*)
uAcc := 16#0000_0000;

IF nCount < nLenUse THEN
    nUse := nCount;             // 不足：只组前 nUse 字节，高段零 / Short: assemble what we have
    uInfoId := 16#0001_04B8;    // 信息级：源字节不足补零 / Info: padded with zeros
ELSE
    nUse := nLenUse;            // 充足：全量组装 / Full assembly
END_IF

FOR i := 0 TO (nUse - 1) DO
    (* 槽位映射（对合映射，与 WordToBytes 同口径，round-trip 成立） *)
    (* Slot mapping, involutive, shared with WordToBytes for round-trip *)
    IF eOrder = E_DL_ByteOrder.eDcba THEN
        nSlot := (nLenUse - 1) - i;          // 全反序 / Full reverse
    ELSIF eOrder = E_DL_ByteOrder.eBadc THEN
        nSlot := (i XOR 1) MOD nLenUse;      // 寄存器内两两互换 / Swap within register pairs
    ELSIF eOrder = E_DL_ByteOrder.eCdab THEN
        IF nLenUse = DL_WFB_LEN_MAX THEN
            nSlot := (i XOR 2) MOD nLenUse;  // DWORD：高低字互换 / DWORD: word swap
        ELSE
            nSlot := 1 - i;                  // WORD：退化为字节反序（见头披露）/ WORD: degenerate reverse
        END_IF
    ELSE
        nSlot := i;                          // eAbcd 大端直排（含越界回退默认）/ Big endian, incl. fallback
    END_IF

    uB     := pBytes[i];                       // 取源字节（指针下标访问）/ Fetch source byte
    nShift := (nLenUse - 1 - nSlot) * 8;       // 槽位移位量 [bit]，DINT 承载，结构性 <= 24 / Slot shift
    uAcc   := uAcc OR SHL(BYTE_TO_DWORD(uB), nShift);    // 升位左移按位或 / Widen, shift, OR
END_FOR

(*------------------------------------------------------------------------------
 * 段 4｜结果回写：WORD 目标结果天然落在低 16 位（槽位 0..1 移位量 0/8），无需再掩码
 *      Result write-back: WORD target lands in the low word by construction
 *-----------------------------------------------------------------------------*)
FC_DL_WordFromBytes := uAcc;
bValid := TRUE;
END_FUNCTION

(* ---- FC_DL_WordToBinString.st ---- *)
(*
    FC_DL_WordToBinString —— WORD → 16 字符定长二进制文本（MSB-first）
    ------------------------------------------------------------------
    组件名称  : FC_DL_WordToBinString
    分类      : DL_MathData / BitText
    前缀      : FC_DL_
    版本      : 1.0.0
    溯源      : IEC 61131-3 标准语义的道莅防御性实现（WORD 位序 → '0'/'1'
                文本化的位掩码提取，与库内 FC_DL_DwordToHexString（十六进制
                文本化）同族反向补口）；实现 / 引脚名 / 码位 100% 自有；
                clean-room 声明 —— 零代码行复制，无闭源参考。
    平台      : 纯 IEC 61131-3（FOR + SHL + CONCAT），无内建函数依赖，
                CODESYS 3.5 / TwinCAT 3 / InoProShop / Machine Expert 通用
    作者      : 道莅代码库 · PLC编程专家（R72 构建轮 · 批 2 · 序号 5）
    ------------------------------------------------------------------
    功能说明  : 把 WORD 的 16 个位按 **MSB-first**（位 15 → 位 0）顺序拼接为
                16 字符定长二进制文本（'0101…'，字符 '1' = 位 1，'0' = 位 0）。
                真实工况：调试面板位诊断显示、协议帧人读文本、培训 / 文档
                向量打印。
                判据链：逐位提取（掩码法：uMask := SHL(WORD#1, uBit)，uBit 由
                常量界循环 0..15 生成，**全程无 64 位移位、移位量 ≤ 15 <
                WORD 位宽 16**（R48 移位量归一：结构性保证，非变量依赖））
                → 定长出口（16 字符恒定，无截断可能——与可截断族的口径差异：
                本件输出长度是输入位宽的常量函数，不随值变化）。
                位序口径声明：MSB-first（位 15 在串首），与网络字节序调试
                惯例一致；LSB-first 需求属另一语义（位序重排归
                FC_DL_ReverseBitsWord，不在本件）。
    错误码    : N/A —— 本件为全定义域全值函数（65536 个 WORD 值全部得到
                确定 16 字符输出），bValid 恒 TRUE 仅保留契约一致性，无故障 /
                信息出口，无码位分配。
    码位总账  : 无（全值函数）
    状态机    : N/A —— 纯函数无状态，无 CASE 可写，非法状态不可能出现
    边界与披露: 一 无定时器 / 无沿检测实例 / 无除法，FOR 循环界为常量
                   0..15（无变量界，无死循环面，守卫计数器豁免），周期安全
                   规则 N/A；
                二 零全局变量、零 VAR_EXTERNAL、零物理地址；
                三 验收向量：V1 uWord = 16#0000 → '0000000000000000'（全 0 串）；
                   V2 uWord = 16#FFFF → '1111111111111111'（全 1 串）；
                   V3 uWord = 16#0001 → '0000000000000001'（LSB 在串尾，
                   MSB-first 口径自证）；V4 uWord = 16#8000 → '1000000000000000'。
                算法已证（脚本）：未跑 ｜ 编译器已证（三平台）：未跑
    分工声明  : FC_DL_DwordToHexString（十六进制文本化）、FC_DL_ReverseBitsWord
                （位序重排非文本化）、FC_DL_FirstSetBit（位搜索）——本件只做
                WORD 的二进制文本化，三者均不替代本件。
    修订记录  : 2026-11-23 v1.0.0 首次入库（R72 构建轮 · 批 2 · 序号 5）
*)
FUNCTION FC_DL_WordToBinString : STRING
VAR_INPUT
    uWord : WORD;                          (* 待文本化字，[位图]，本件不解释位语义 / the word under conversion, the FC never interprets bit semantics *)
END_VAR
VAR_OUTPUT
    bValid : BOOL;                         (* 输出可用标志，恒 TRUE（契约一致性保留）/ the outputs usable flag, always TRUE by contract *)
END_VAR
VAR CONSTANT
    DL_WBS_ONE   : STRING(1) := '1';       // 位 1 字符 [文本] / the bit one char
    DL_WBS_ZERO  : STRING(1) := '0';       // 位 0 字符 [文本] / the bit zero char
    DL_WBS_BITS  : INT := 16;              (* WORD 位宽（常量界循环上界 − 1）[位] / the word width *)
    DL_WBS_LAST  : INT := 15;              (* MSB-first 首位下标（位 15）[位] / the first bit index, MSB first *)
    DL_WBS_STEP  : INT := 1;               (* 循环步进 [位] / the loop step *)
    DL_WBS_ZEROI : INT := 0;               (* LSB 循环下界 [位] / the loop lower bound *)
END_VAR
VAR
    nI    : INT;                           (* 循环游标（0..15，常量界）[位] / the loop cursor *)
    uBit  : INT;                           (* 当前提取位号（15 − nI，MSB-first）[位] / the current bit index *)
    uMask : WORD;                          (* 当前位掩码 [位图] / the current bit mask *)
END_VAR

// 段 1｜返回值与状态预置（统一出口预置，R256）/ segment 1, preset the return and the status
FC_DL_WordToBinString := '';             // 预置空串，逐位拼接 / preset the empty string
bValid := FALSE;                         // 预置不可用，出口翻转 / preset unusable
nI    := DL_WBS_ZEROI;                   // 游标预置 / preset the cursor
uBit  := DL_WBS_LAST;                    // 位号预置（MSB-first 起点）/ preset the bit index
uMask := WORD#0;                         // 掩码清零 / clear the mask

// 段 2｜逐位提取拼接（位 15 → 位 0，MSB-first；移位量 uBit ∈ [0,15] 结构性
//        小于位宽 16，R48 归一豁免声明）/ segment 2, the bit by bit extraction
FOR nI := DL_WBS_ZEROI TO DL_WBS_LAST BY DL_WBS_STEP DO // 常量界循环（无变量界死循环面）/ the constant bound loop
    uBit := DL_WBS_LAST - nI;            // MSB-first 位号 / the MSB first bit index
    uMask := SHL(WORD#1, uBit);          // 掩码法取位（移位量 <= 15，结构性安全）/ the mask method
    IF (uWord AND uMask) <> WORD#0 THEN  // 位为 1 / the bit is one
        FC_DL_WordToBinString := CONCAT(FC_DL_WordToBinString, DL_WBS_ONE); // 拼 '1' / append the one char
    ELSE                                 // 位为 0 / the bit is zero
        FC_DL_WordToBinString := CONCAT(FC_DL_WordToBinString, DL_WBS_ZERO); // 拼 '0' / append the zero char
    END_IF
END_FOR

// 段 3｜统一出口（16 字符恒定，无截断可能）/ segment 3, the unified outlet
bValid := TRUE;                          // 全值函数恒可用 / the total function always usable
END_FUNCTION
